DATA_BLOCK "TCP_IP_Shuttle_DB_20"   // DB238
{ S7_Optimized_Access := 'TRUE' }
VERSION : 0.1
// stored: AutoNumber true, DBAccessibleFromOPCUA true, IsOnlyStoredInLoadMemory false, IsRetainMemResEnabled false, IsWriteProtectedInAS false, MemoryReserve 100
   VAR
      enable : Bool := TRUE;
      send : Bool;
      sendDataLength : UDInt := 0;
      receiveDataLength : UDInt := 16#FFFF_FFFF;
   END_VAR
   VAR RETAIN
      tcpConfig : "LCom_typeConfig";
   END_VAR
   VAR
      tcpDiagnostics { S7_SetPoint := 'True'} : "LCom_typeDiagnostics";
      sendBuffer { S7_SetPoint := 'True'} : Array[0..59] of Byte;
      SendBufferSize : UInt := 60;
      receiveBuffer : Array[0..27] of Byte;
      receiveBufferSize : UInt := 28;
      connected : Bool;
      sending : Bool;
      dataReceived : Bool;
      receivedDataLength : UDInt;
      busy : Bool;
      error : Bool;
      status : Word;
   END_VAR
BEGIN
   tcpConfig.connection.interfaceID := 65164;
   tcpConfig.connection.connectionID := 120;
   tcpConfig.connection.comService := 1;
   tcpConfig.connection.isClient := False;
   tcpConfig.connection.connectType := 1;
   tcpConfig.connection.localPort := 4020;
   tcpConfig.connection.partnerPort := 4020;
   tcpConfig.connection.partnerIP.ADDR[1] := 10;
   tcpConfig.connection.partnerIP.ADDR[2] := 0;
   tcpConfig.connection.partnerIP.ADDR[3] := 34;
   tcpConfig.connection.partnerIP.ADDR[4] := 230;
   tcpConfig.connection.acceptUnknownPartner := TRUE;
   tcpConfig.connection.lifeSignCycleTime := T#1s;
   // sendBuffer[0] : STX
   // sendBuffer[1] : Size
   // sendBuffer[2] : Type
   // sendBuffer[3] : Request ID 1
   // sendBuffer[4] : Request ID 2
   // sendBuffer[5] : PID 1
   // sendBuffer[6] : PID 2
   // sendBuffer[7] : PID 3
   // sendBuffer[8] : PID 4
   // sendBuffer[9] : DID 1
   // sendBuffer[10] : DID 2
   // sendBuffer[11] : DID 3
   // sendBuffer[12] : DID 4
   // sendBuffer[13] : Distance remaining 1
   // sendBuffer[14] : Distance remaining 2
   // sendBuffer[15] : X
   // sendBuffer[16] : X
   // sendBuffer[17] : X
   // sendBuffer[18] : X
   // sendBuffer[19] : Y
   // sendBuffer[20] : Y
   // sendBuffer[21] : Y
   // sendBuffer[22] : Y
   // sendBuffer[23] : Floor
   // sendBuffer[24] : Mode
   // sendBuffer[25] : State
   // sendBuffer[26] : Load State
   // sendBuffer[27] : E1
   // sendBuffer[28] : E1
   // sendBuffer[29] : E2
   // sendBuffer[30] : E2
   // sendBuffer[31] : E3
   // sendBuffer[32] : E3
   // sendBuffer[33] : E4
   // sendBuffer[34] : E4
   // sendBuffer[35] : E5
   // sendBuffer[36] : E5
   // sendBuffer[37] : E6
   // sendBuffer[38] : E6
   // sendBuffer[39] : I1
   // sendBuffer[40] : I1
   // sendBuffer[41] : Q1
   // sendBuffer[42] : Q1
   // sendBuffer[43] : Barcode 1
   // sendBuffer[44] : Barcode 2
   // sendBuffer[45] : Barcode 3
   // sendBuffer[46] : Barcode 4
   // sendBuffer[47] : Pallet Type
   // sendBuffer[48] : Energy Level
   // sendBuffer[49] : Battery Voltage
   // sendBuffer[50] : Battery Voltage
   // sendBuffer[51] : Paused
   // sendBuffer[52] : Last order 1
   // sendBuffer[53] : Last order 2
   // sendBuffer[54] : Current order 1
   // sendBuffer[55] : Current order 2
   // sendBuffer[56] : Last finished 1
   // sendBuffer[57] : Last Finished 2
   // sendBuffer[58] : CS
   // sendBuffer[59] : ETX
   // receiveBuffer[0] : STX
   // receiveBuffer[1] : Size (length of payload)
   // receiveBuffer[2] : Type
   // receiveBuffer[3] : Request ID 1
   // receiveBuffer[4] : Request ID 2
END_DATA_BLOCK

DATA_BLOCK "TCP_IP_Shuttle_DB_21"   // DB166
{ S7_Optimized_Access := 'TRUE' }
VERSION : 0.1
// stored: AutoNumber true, DBAccessibleFromOPCUA true, IsOnlyStoredInLoadMemory false, IsRetainMemResEnabled false, IsWriteProtectedInAS false, MemoryReserve 100
   VAR
      enable : Bool := TRUE;
      send : Bool;
      sendDataLength : UDInt := 0;
      receiveDataLength : UDInt := 16#FFFF_FFFF;
   END_VAR
   VAR RETAIN
      tcpConfig : "LCom_typeConfig";
   END_VAR
   VAR
      tcpDiagnostics { S7_SetPoint := 'True'} : "LCom_typeDiagnostics";
      sendBuffer { S7_SetPoint := 'True'} : Array[0..59] of Byte;
      SendBufferSize : UInt := 60;
      receiveBuffer : Array[0..27] of Byte;
      receiveBufferSize : UInt := 28;
      connected : Bool;
      sending : Bool;
      dataReceived : Bool;
      receivedDataLength : UDInt;
      busy : Bool;
      error : Bool;
      status : Word;
   END_VAR
BEGIN
   tcpConfig.connection.interfaceID := 65164;
   tcpConfig.connection.connectionID := 121;
   tcpConfig.connection.comService := 1;
   tcpConfig.connection.isClient := False;
   tcpConfig.connection.connectType := 1;
   tcpConfig.connection.localPort := 4021;
   tcpConfig.connection.partnerPort := 4021;
   tcpConfig.connection.partnerIP.ADDR[1] := 10;
   tcpConfig.connection.partnerIP.ADDR[2] := 0;
   tcpConfig.connection.partnerIP.ADDR[3] := 34;
   tcpConfig.connection.partnerIP.ADDR[4] := 231;
   tcpConfig.connection.acceptUnknownPartner := TRUE;
   tcpConfig.connection.lifeSignCycleTime := T#1s;
   // sendBuffer[0] : STX
   // sendBuffer[1] : Size
   // sendBuffer[2] : Type
   // sendBuffer[3] : Request ID 1
   // sendBuffer[4] : Request ID 2
   // sendBuffer[5] : PID 1
   // sendBuffer[6] : PID 2
   // sendBuffer[7] : PID 3
   // sendBuffer[8] : PID 4
   // sendBuffer[9] : DID 1
   // sendBuffer[10] : DID 2
   // sendBuffer[11] : DID 3
   // sendBuffer[12] : DID 4
   // sendBuffer[13] : Distance remaining 1
   // sendBuffer[14] : Distance remaining 2
   // sendBuffer[15] : X
   // sendBuffer[16] : X
   // sendBuffer[17] : X
   // sendBuffer[18] : X
   // sendBuffer[19] : Y
   // sendBuffer[20] : Y
   // sendBuffer[21] : Y
   // sendBuffer[22] : Y
   // sendBuffer[23] : Floor
   // sendBuffer[24] : Mode
   // sendBuffer[25] : State
   // sendBuffer[26] : Load State
   // sendBuffer[27] : E1
   // sendBuffer[28] : E1
   // sendBuffer[29] : E2
   // sendBuffer[30] : E2
   // sendBuffer[31] : E3
   // sendBuffer[32] : E3
   // sendBuffer[33] : E4
   // sendBuffer[34] : E4
   // sendBuffer[35] : E5
   // sendBuffer[36] : E5
   // sendBuffer[37] : E6
   // sendBuffer[38] : E6
   // sendBuffer[39] : I1
   // sendBuffer[40] : I1
   // sendBuffer[41] : Q1
   // sendBuffer[42] : Q1
   // sendBuffer[43] : Barcode 1
   // sendBuffer[44] : Barcode 2
   // sendBuffer[45] : Barcode 3
   // sendBuffer[46] : Barcode 4
   // sendBuffer[47] : Pallet Type
   // sendBuffer[48] : Energy Level
   // sendBuffer[49] : Battery Voltage
   // sendBuffer[50] : Battery Voltage
   // sendBuffer[51] : Paused
   // sendBuffer[52] : Last order 1
   // sendBuffer[53] : Last order 2
   // sendBuffer[54] : Current order 1
   // sendBuffer[55] : Current order 2
   // sendBuffer[56] : Last finished 1
   // sendBuffer[57] : Last Finished 2
   // sendBuffer[58] : CS
   // sendBuffer[59] : ETX
   // receiveBuffer[0] : STX
   // receiveBuffer[1] : Size (length of payload)
   // receiveBuffer[2] : Type
   // receiveBuffer[3] : Request ID 1
   // receiveBuffer[4] : Request ID 2
END_DATA_BLOCK

DATA_BLOCK "TCP_IP_Shuttle_DB_22"   // DB241
{ S7_Optimized_Access := 'TRUE' }
VERSION : 0.1
// stored: AutoNumber true, DBAccessibleFromOPCUA true, IsOnlyStoredInLoadMemory false, IsRetainMemResEnabled false, IsWriteProtectedInAS false, MemoryReserve 100
   VAR
      enable : Bool := TRUE;
      send : Bool;
      sendDataLength : UDInt := 0;
      receiveDataLength : UDInt := 16#FFFF_FFFF;
   END_VAR
   VAR RETAIN
      tcpConfig : "LCom_typeConfig";
   END_VAR
   VAR
      tcpDiagnostics { S7_SetPoint := 'True'} : "LCom_typeDiagnostics";
      sendBuffer { S7_SetPoint := 'True'} : Array[0..59] of Byte;
      SendBufferSize : UInt := 60;
      receiveBuffer : Array[0..27] of Byte;
      receiveBufferSize : UInt := 28;
      connected : Bool;
      sending : Bool;
      dataReceived : Bool;
      receivedDataLength : UDInt;
      busy : Bool;
      error : Bool;
      status : Word;
   END_VAR
BEGIN
   tcpConfig.connection.interfaceID := 65164;
   tcpConfig.connection.connectionID := 122;
   tcpConfig.connection.comService := 1;
   tcpConfig.connection.isClient := False;
   tcpConfig.connection.connectType := 1;
   tcpConfig.connection.localPort := 4022;
   tcpConfig.connection.partnerPort := 4022;
   tcpConfig.connection.partnerIP.ADDR[1] := 10;
   tcpConfig.connection.partnerIP.ADDR[2] := 0;
   tcpConfig.connection.partnerIP.ADDR[3] := 34;
   tcpConfig.connection.partnerIP.ADDR[4] := 232;
   tcpConfig.connection.acceptUnknownPartner := TRUE;
   tcpConfig.connection.lifeSignCycleTime := T#1s;
   // sendBuffer[0] : STX
   // sendBuffer[1] : Size
   // sendBuffer[2] : Type
   // sendBuffer[3] : Request ID 1
   // sendBuffer[4] : Request ID 2
   // sendBuffer[5] : PID 1
   // sendBuffer[6] : PID 2
   // sendBuffer[7] : PID 3
   // sendBuffer[8] : PID 4
   // sendBuffer[9] : DID 1
   // sendBuffer[10] : DID 2
   // sendBuffer[11] : DID 3
   // sendBuffer[12] : DID 4
   // sendBuffer[13] : Distance remaining 1
   // sendBuffer[14] : Distance remaining 2
   // sendBuffer[15] : X
   // sendBuffer[16] : X
   // sendBuffer[17] : X
   // sendBuffer[18] : X
   // sendBuffer[19] : Y
   // sendBuffer[20] : Y
   // sendBuffer[21] : Y
   // sendBuffer[22] : Y
   // sendBuffer[23] : Floor
   // sendBuffer[24] : Mode
   // sendBuffer[25] : State
   // sendBuffer[26] : Load State
   // sendBuffer[27] : E1
   // sendBuffer[28] : E1
   // sendBuffer[29] : E2
   // sendBuffer[30] : E2
   // sendBuffer[31] : E3
   // sendBuffer[32] : E3
   // sendBuffer[33] : E4
   // sendBuffer[34] : E4
   // sendBuffer[35] : E5
   // sendBuffer[36] : E5
   // sendBuffer[37] : E6
   // sendBuffer[38] : E6
   // sendBuffer[39] : I1
   // sendBuffer[40] : I1
   // sendBuffer[41] : Q1
   // sendBuffer[42] : Q1
   // sendBuffer[43] : Barcode 1
   // sendBuffer[44] : Barcode 2
   // sendBuffer[45] : Barcode 3
   // sendBuffer[46] : Barcode 4
   // sendBuffer[47] : Pallet Type
   // sendBuffer[48] : Energy Level
   // sendBuffer[49] : Battery Voltage
   // sendBuffer[50] : Battery Voltage
   // sendBuffer[51] : Paused
   // sendBuffer[52] : Last order 1
   // sendBuffer[53] : Last order 2
   // sendBuffer[54] : Current order 1
   // sendBuffer[55] : Current order 2
   // sendBuffer[56] : Last finished 1
   // sendBuffer[57] : Last Finished 2
   // sendBuffer[58] : CS
   // sendBuffer[59] : ETX
   // receiveBuffer[0] : STX
   // receiveBuffer[1] : Size (length of payload)
   // receiveBuffer[2] : Type
   // receiveBuffer[3] : Request ID 1
   // receiveBuffer[4] : Request ID 2
END_DATA_BLOCK

DATA_BLOCK "TCP_IP_Shuttle_DB_23"   // DB382
{ S7_Optimized_Access := 'TRUE' }
VERSION : 0.1
// stored: AutoNumber true, DBAccessibleFromOPCUA true, IsOnlyStoredInLoadMemory false, IsRetainMemResEnabled false, IsWriteProtectedInAS false, MemoryReserve 100
   VAR
      enable : Bool := TRUE;
      send : Bool;
      sendDataLength : UDInt := 0;
      receiveDataLength : UDInt := 16#FFFF_FFFF;
   END_VAR
   VAR RETAIN
      tcpConfig : "LCom_typeConfig";
   END_VAR
   VAR
      tcpDiagnostics { S7_SetPoint := 'True'} : "LCom_typeDiagnostics";
      sendBuffer { S7_SetPoint := 'True'} : Array[0..59] of Byte;
      SendBufferSize : UInt := 60;
      receiveBuffer : Array[0..27] of Byte;
      receiveBufferSize : UInt := 28;
      connected : Bool;
      sending : Bool;
      dataReceived : Bool;
      receivedDataLength : UDInt;
      busy : Bool;
      error : Bool;
      status : Word;
   END_VAR
BEGIN
   tcpConfig.connection.interfaceID := 65164;
   tcpConfig.connection.connectionID := 123;
   tcpConfig.connection.comService := 1;
   tcpConfig.connection.isClient := False;
   tcpConfig.connection.connectType := 1;
   tcpConfig.connection.localPort := 4023;
   tcpConfig.connection.partnerPort := 4023;
   tcpConfig.connection.partnerIP.ADDR[1] := 10;
   tcpConfig.connection.partnerIP.ADDR[2] := 0;
   tcpConfig.connection.partnerIP.ADDR[3] := 34;
   tcpConfig.connection.partnerIP.ADDR[4] := 233;
   tcpConfig.connection.acceptUnknownPartner := TRUE;
   tcpConfig.connection.lifeSignCycleTime := T#1s;
   // sendBuffer[0] : STX
   // sendBuffer[1] : Size
   // sendBuffer[2] : Type
   // sendBuffer[3] : Request ID 1
   // sendBuffer[4] : Request ID 2
   // sendBuffer[5] : PID 1
   // sendBuffer[6] : PID 2
   // sendBuffer[7] : PID 3
   // sendBuffer[8] : PID 4
   // sendBuffer[9] : DID 1
   // sendBuffer[10] : DID 2
   // sendBuffer[11] : DID 3
   // sendBuffer[12] : DID 4
   // sendBuffer[13] : Distance remaining 1
   // sendBuffer[14] : Distance remaining 2
   // sendBuffer[15] : X
   // sendBuffer[16] : X
   // sendBuffer[17] : X
   // sendBuffer[18] : X
   // sendBuffer[19] : Y
   // sendBuffer[20] : Y
   // sendBuffer[21] : Y
   // sendBuffer[22] : Y
   // sendBuffer[23] : Floor
   // sendBuffer[24] : Mode
   // sendBuffer[25] : State
   // sendBuffer[26] : Load State
   // sendBuffer[27] : E1
   // sendBuffer[28] : E1
   // sendBuffer[29] : E2
   // sendBuffer[30] : E2
   // sendBuffer[31] : E3
   // sendBuffer[32] : E3
   // sendBuffer[33] : E4
   // sendBuffer[34] : E4
   // sendBuffer[35] : E5
   // sendBuffer[36] : E5
   // sendBuffer[37] : E6
   // sendBuffer[38] : E6
   // sendBuffer[39] : I1
   // sendBuffer[40] : I1
   // sendBuffer[41] : Q1
   // sendBuffer[42] : Q1
   // sendBuffer[43] : Barcode 1
   // sendBuffer[44] : Barcode 2
   // sendBuffer[45] : Barcode 3
   // sendBuffer[46] : Barcode 4
   // sendBuffer[47] : Pallet Type
   // sendBuffer[48] : Energy Level
   // sendBuffer[49] : Battery Voltage
   // sendBuffer[50] : Battery Voltage
   // sendBuffer[51] : Paused
   // sendBuffer[52] : Last order 1
   // sendBuffer[53] : Last order 2
   // sendBuffer[54] : Current order 1
   // sendBuffer[55] : Current order 2
   // sendBuffer[56] : Last finished 1
   // sendBuffer[57] : Last Finished 2
   // sendBuffer[58] : CS
   // sendBuffer[59] : ETX
   // receiveBuffer[0] : STX
   // receiveBuffer[1] : Size (length of payload)
   // receiveBuffer[2] : Type
   // receiveBuffer[3] : Request ID 1
   // receiveBuffer[4] : Request ID 2
END_DATA_BLOCK

DATA_BLOCK "TCP_IP_Shuttle_DB_3"   // DB388
{ S7_Optimized_Access := 'TRUE' }
VERSION : 0.1
// stored: AutoNumber true, DBAccessibleFromOPCUA true, IsOnlyStoredInLoadMemory false, IsRetainMemResEnabled false, IsWriteProtectedInAS false, MemoryReserve 100
   VAR
      enable : Bool := TRUE;
      send : Bool;
      sendDataLength : UDInt := 0;
      receiveDataLength : UDInt := 16#FFFF_FFFF;
   END_VAR
   VAR RETAIN
      tcpConfig : "LCom_typeConfig";
   END_VAR
   VAR
      tcpDiagnostics { S7_SetPoint := 'True'} : "LCom_typeDiagnostics";
      sendBuffer { S7_SetPoint := 'True'} : Array[0..59] of Byte;
      SendBufferSize : UInt := 60;
      receiveBuffer : Array[0..27] of Byte;
      receiveBufferSize : UInt := 28;
      connected : Bool;
      sending : Bool;
      dataReceived : Bool;
      receivedDataLength : UDInt;
      busy : Bool;
      error : Bool;
      status : Word;
   END_VAR
BEGIN
   tcpConfig.connection.interfaceID := 65164;
   tcpConfig.connection.connectionID := 103;
   tcpConfig.connection.comService := 1;
   tcpConfig.connection.isClient := False;
   tcpConfig.connection.connectType := 1;
   tcpConfig.connection.localPort := 4003;
   tcpConfig.connection.partnerPort := 4003;
   tcpConfig.connection.partnerIP.ADDR[1] := 10;
   tcpConfig.connection.partnerIP.ADDR[2] := 0;
   tcpConfig.connection.partnerIP.ADDR[3] := 34;
   tcpConfig.connection.partnerIP.ADDR[4] := 213;
   tcpConfig.connection.acceptUnknownPartner := TRUE;
   tcpConfig.connection.lifeSignCycleTime := T#1s;
   // sendBuffer[0] : STX
   // sendBuffer[1] : Size
   // sendBuffer[2] : Type
   // sendBuffer[3] : Request ID 1
   // sendBuffer[4] : Request ID 2
   // sendBuffer[5] : PID 1
   // sendBuffer[6] : PID 2
   // sendBuffer[7] : PID 3
   // sendBuffer[8] : PID 4
   // sendBuffer[9] : DID 1
   // sendBuffer[10] : DID 2
   // sendBuffer[11] : DID 3
   // sendBuffer[12] : DID 4
   // sendBuffer[13] : Distance remaining 1
   // sendBuffer[14] : Distance remaining 2
   // sendBuffer[15] : X
   // sendBuffer[16] : X
   // sendBuffer[17] : X
   // sendBuffer[18] : X
   // sendBuffer[19] : Y
   // sendBuffer[20] : Y
   // sendBuffer[21] : Y
   // sendBuffer[22] : Y
   // sendBuffer[23] : Floor
   // sendBuffer[24] : Mode
   // sendBuffer[25] : State
   // sendBuffer[26] : Load State
   // sendBuffer[27] : E1
   // sendBuffer[28] : E1
   // sendBuffer[29] : E2
   // sendBuffer[30] : E2
   // sendBuffer[31] : E3
   // sendBuffer[32] : E3
   // sendBuffer[33] : E4
   // sendBuffer[34] : E4
   // sendBuffer[35] : E5
   // sendBuffer[36] : E5
   // sendBuffer[37] : E6
   // sendBuffer[38] : E6
   // sendBuffer[39] : I1
   // sendBuffer[40] : I1
   // sendBuffer[41] : Q1
   // sendBuffer[42] : Q1
   // sendBuffer[43] : Barcode 1
   // sendBuffer[44] : Barcode 2
   // sendBuffer[45] : Barcode 3
   // sendBuffer[46] : Barcode 4
   // sendBuffer[47] : Pallet Type
   // sendBuffer[48] : Energy Level
   // sendBuffer[49] : Battery Voltage
   // sendBuffer[50] : Battery Voltage
   // sendBuffer[51] : Paused
   // sendBuffer[52] : Last order 1
   // sendBuffer[53] : Last order 2
   // sendBuffer[54] : Current order 1
   // sendBuffer[55] : Current order 2
   // sendBuffer[56] : Last finished 1
   // sendBuffer[57] : Last Finished 2
   // sendBuffer[58] : CS
   // sendBuffer[59] : ETX
   // receiveBuffer[0] : STX
   // receiveBuffer[1] : Size (length of payload)
   // receiveBuffer[2] : Type
   // receiveBuffer[3] : Request ID 1
   // receiveBuffer[4] : Request ID 2
END_DATA_BLOCK

DATA_BLOCK "TCP_IP_Shuttle_DB_4"   // DB375
{ S7_Optimized_Access := 'TRUE' }
VERSION : 0.1
// stored: AutoNumber true, DBAccessibleFromOPCUA true, IsOnlyStoredInLoadMemory false, IsRetainMemResEnabled false, IsWriteProtectedInAS false, MemoryReserve 100
   VAR
      enable : Bool := TRUE;
      send : Bool;
      sendDataLength : UDInt := 0;
      receiveDataLength : UDInt := 16#FFFF_FFFF;
   END_VAR
   VAR RETAIN
      tcpConfig : "LCom_typeConfig";
   END_VAR
   VAR
      tcpDiagnostics { S7_SetPoint := 'True'} : "LCom_typeDiagnostics";
      sendBuffer { S7_SetPoint := 'True'} : Array[0..59] of Byte;
      SendBufferSize : UInt := 60;
      receiveBuffer : Array[0..27] of Byte;
      receiveBufferSize : UInt := 28;
      connected : Bool;
      sending : Bool;
      dataReceived : Bool;
      receivedDataLength : UDInt;
      busy : Bool;
      error : Bool;
      status : Word;
   END_VAR
BEGIN
   tcpConfig.connection.interfaceID := 65164;
   tcpConfig.connection.connectionID := 104;
   tcpConfig.connection.comService := 1;
   tcpConfig.connection.isClient := False;
   tcpConfig.connection.connectType := 1;
   tcpConfig.connection.localPort := 4004;
   tcpConfig.connection.partnerPort := 4004;
   tcpConfig.connection.partnerIP.ADDR[1] := 10;
   tcpConfig.connection.partnerIP.ADDR[2] := 0;
   tcpConfig.connection.partnerIP.ADDR[3] := 34;
   tcpConfig.connection.partnerIP.ADDR[4] := 214;
   tcpConfig.connection.acceptUnknownPartner := TRUE;
   tcpConfig.connection.lifeSignCycleTime := T#1s;
   // sendBuffer[0] : STX
   // sendBuffer[1] : Size
   // sendBuffer[2] : Type
   // sendBuffer[3] : Request ID 1
   // sendBuffer[4] : Request ID 2
   // sendBuffer[5] : PID 1
   // sendBuffer[6] : PID 2
   // sendBuffer[7] : PID 3
   // sendBuffer[8] : PID 4
   // sendBuffer[9] : DID 1
   // sendBuffer[10] : DID 2
   // sendBuffer[11] : DID 3
   // sendBuffer[12] : DID 4
   // sendBuffer[13] : Distance remaining 1
   // sendBuffer[14] : Distance remaining 2
   // sendBuffer[15] : X
   // sendBuffer[16] : X
   // sendBuffer[17] : X
   // sendBuffer[18] : X
   // sendBuffer[19] : Y
   // sendBuffer[20] : Y
   // sendBuffer[21] : Y
   // sendBuffer[22] : Y
   // sendBuffer[23] : Floor
   // sendBuffer[24] : Mode
   // sendBuffer[25] : State
   // sendBuffer[26] : Load State
   // sendBuffer[27] : E1
   // sendBuffer[28] : E1
   // sendBuffer[29] : E2
   // sendBuffer[30] : E2
   // sendBuffer[31] : E3
   // sendBuffer[32] : E3
   // sendBuffer[33] : E4
   // sendBuffer[34] : E4
   // sendBuffer[35] : E5
   // sendBuffer[36] : E5
   // sendBuffer[37] : E6
   // sendBuffer[38] : E6
   // sendBuffer[39] : I1
   // sendBuffer[40] : I1
   // sendBuffer[41] : Q1
   // sendBuffer[42] : Q1
   // sendBuffer[43] : Barcode 1
   // sendBuffer[44] : Barcode 2
   // sendBuffer[45] : Barcode 3
   // sendBuffer[46] : Barcode 4
   // sendBuffer[47] : Pallet Type
   // sendBuffer[48] : Energy Level
   // sendBuffer[49] : Battery Voltage
   // sendBuffer[50] : Battery Voltage
   // sendBuffer[51] : Paused
   // sendBuffer[52] : Last order 1
   // sendBuffer[53] : Last order 2
   // sendBuffer[54] : Current order 1
   // sendBuffer[55] : Current order 2
   // sendBuffer[56] : Last finished 1
   // sendBuffer[57] : Last Finished 2
   // sendBuffer[58] : CS
   // sendBuffer[59] : ETX
   // receiveBuffer[0] : STX
   // receiveBuffer[1] : Size (length of payload)
   // receiveBuffer[2] : Type
   // receiveBuffer[3] : Request ID 1
   // receiveBuffer[4] : Request ID 2
END_DATA_BLOCK

DATA_BLOCK "TCP_IP_Shuttle_DB_5"   // DB376
{ S7_Optimized_Access := 'TRUE' }
VERSION : 0.1
// stored: AutoNumber true, DBAccessibleFromOPCUA true, IsOnlyStoredInLoadMemory false, IsRetainMemResEnabled false, IsWriteProtectedInAS false, MemoryReserve 100
   VAR
      enable : Bool := TRUE;
      send : Bool;
      sendDataLength : UDInt := 0;
      receiveDataLength : UDInt := 16#FFFF_FFFF;
   END_VAR
   VAR RETAIN
      tcpConfig : "LCom_typeConfig";
   END_VAR
   VAR
      tcpDiagnostics { S7_SetPoint := 'True'} : "LCom_typeDiagnostics";
      sendBuffer { S7_SetPoint := 'True'} : Array[0..59] of Byte;
      SendBufferSize : UInt := 60;
      receiveBuffer : Array[0..27] of Byte;
      receiveBufferSize : UInt := 28;
      connected : Bool;
      sending : Bool;
      dataReceived : Bool;
      receivedDataLength : UDInt;
      busy : Bool;
      error : Bool;
      status : Word;
   END_VAR
BEGIN
   tcpConfig.connection.interfaceID := 65164;
   tcpConfig.connection.connectionID := 105;
   tcpConfig.connection.comService := 1;
   tcpConfig.connection.isClient := False;
   tcpConfig.connection.connectType := 1;
   tcpConfig.connection.localPort := 4005;
   tcpConfig.connection.partnerPort := 4005;
   tcpConfig.connection.partnerIP.ADDR[1] := 10;
   tcpConfig.connection.partnerIP.ADDR[2] := 0;
   tcpConfig.connection.partnerIP.ADDR[3] := 34;
   tcpConfig.connection.partnerIP.ADDR[4] := 215;
   tcpConfig.connection.acceptUnknownPartner := TRUE;
   tcpConfig.connection.lifeSignCycleTime := T#1s;
   // sendBuffer[0] : STX
   // sendBuffer[1] : Size
   // sendBuffer[2] : Type
   // sendBuffer[3] : Request ID 1
   // sendBuffer[4] : Request ID 2
   // sendBuffer[5] : PID 1
   // sendBuffer[6] : PID 2
   // sendBuffer[7] : PID 3
   // sendBuffer[8] : PID 4
   // sendBuffer[9] : DID 1
   // sendBuffer[10] : DID 2
   // sendBuffer[11] : DID 3
   // sendBuffer[12] : DID 4
   // sendBuffer[13] : Distance remaining 1
   // sendBuffer[14] : Distance remaining 2
   // sendBuffer[15] : X
   // sendBuffer[16] : X
   // sendBuffer[17] : X
   // sendBuffer[18] : X
   // sendBuffer[19] : Y
   // sendBuffer[20] : Y
   // sendBuffer[21] : Y
   // sendBuffer[22] : Y
   // sendBuffer[23] : Floor
   // sendBuffer[24] : Mode
   // sendBuffer[25] : State
   // sendBuffer[26] : Load State
   // sendBuffer[27] : E1
   // sendBuffer[28] : E1
   // sendBuffer[29] : E2
   // sendBuffer[30] : E2
   // sendBuffer[31] : E3
   // sendBuffer[32] : E3
   // sendBuffer[33] : E4
   // sendBuffer[34] : E4
   // sendBuffer[35] : E5
   // sendBuffer[36] : E5
   // sendBuffer[37] : E6
   // sendBuffer[38] : E6
   // sendBuffer[39] : I1
   // sendBuffer[40] : I1
   // sendBuffer[41] : Q1
   // sendBuffer[42] : Q1
   // sendBuffer[43] : Barcode 1
   // sendBuffer[44] : Barcode 2
   // sendBuffer[45] : Barcode 3
   // sendBuffer[46] : Barcode 4
   // sendBuffer[47] : Pallet Type
   // sendBuffer[48] : Energy Level
   // sendBuffer[49] : Battery Voltage
   // sendBuffer[50] : Battery Voltage
   // sendBuffer[51] : Paused
   // sendBuffer[52] : Last order 1
   // sendBuffer[53] : Last order 2
   // sendBuffer[54] : Current order 1
   // sendBuffer[55] : Current order 2
   // sendBuffer[56] : Last finished 1
   // sendBuffer[57] : Last Finished 2
   // sendBuffer[58] : CS
   // sendBuffer[59] : ETX
   // receiveBuffer[0] : STX
   // receiveBuffer[1] : Size (length of payload)
   // receiveBuffer[2] : Type
   // receiveBuffer[3] : Request ID 1
   // receiveBuffer[4] : Request ID 2
END_DATA_BLOCK

DATA_BLOCK "TCP_IP_Shuttle_DB_6"   // DB377
{ S7_Optimized_Access := 'TRUE' }
VERSION : 0.1
// stored: AutoNumber true, DBAccessibleFromOPCUA true, IsOnlyStoredInLoadMemory false, IsRetainMemResEnabled false, IsWriteProtectedInAS false, MemoryReserve 100
   VAR
      enable : Bool := TRUE;
      send : Bool;
      sendDataLength : UDInt := 0;
      receiveDataLength : UDInt := 16#FFFF_FFFF;
   END_VAR
   VAR RETAIN
      tcpConfig : "LCom_typeConfig";
   END_VAR
   VAR
      tcpDiagnostics { S7_SetPoint := 'True'} : "LCom_typeDiagnostics";
      sendBuffer { S7_SetPoint := 'True'} : Array[0..59] of Byte;
      SendBufferSize : UInt := 60;
      receiveBuffer : Array[0..27] of Byte;
      receiveBufferSize : UInt := 28;
      connected : Bool;
      sending : Bool;
      dataReceived : Bool;
      receivedDataLength : UDInt;
      busy : Bool;
      error : Bool;
      status : Word;
   END_VAR
BEGIN
   tcpConfig.connection.interfaceID := 65164;
   tcpConfig.connection.connectionID := 106;
   tcpConfig.connection.comService := 1;
   tcpConfig.connection.isClient := False;
   tcpConfig.connection.connectType := 1;
   tcpConfig.connection.localPort := 4006;
   tcpConfig.connection.partnerPort := 4006;
   tcpConfig.connection.partnerIP.ADDR[1] := 10;
   tcpConfig.connection.partnerIP.ADDR[2] := 0;
   tcpConfig.connection.partnerIP.ADDR[3] := 34;
   tcpConfig.connection.partnerIP.ADDR[4] := 216;
   tcpConfig.connection.acceptUnknownPartner := TRUE;
   tcpConfig.connection.lifeSignCycleTime := T#1s;
   // sendBuffer[0] : STX
   // sendBuffer[1] : Size
   // sendBuffer[2] : Type
   // sendBuffer[3] : Request ID 1
   // sendBuffer[4] : Request ID 2
   // sendBuffer[5] : PID 1
   // sendBuffer[6] : PID 2
   // sendBuffer[7] : PID 3
   // sendBuffer[8] : PID 4
   // sendBuffer[9] : DID 1
   // sendBuffer[10] : DID 2
   // sendBuffer[11] : DID 3
   // sendBuffer[12] : DID 4
   // sendBuffer[13] : Distance remaining 1
   // sendBuffer[14] : Distance remaining 2
   // sendBuffer[15] : X
   // sendBuffer[16] : X
   // sendBuffer[17] : X
   // sendBuffer[18] : X
   // sendBuffer[19] : Y
   // sendBuffer[20] : Y
   // sendBuffer[21] : Y
   // sendBuffer[22] : Y
   // sendBuffer[23] : Floor
   // sendBuffer[24] : Mode
   // sendBuffer[25] : State
   // sendBuffer[26] : Load State
   // sendBuffer[27] : E1
   // sendBuffer[28] : E1
   // sendBuffer[29] : E2
   // sendBuffer[30] : E2
   // sendBuffer[31] : E3
   // sendBuffer[32] : E3
   // sendBuffer[33] : E4
   // sendBuffer[34] : E4
   // sendBuffer[35] : E5
   // sendBuffer[36] : E5
   // sendBuffer[37] : E6
   // sendBuffer[38] : E6
   // sendBuffer[39] : I1
   // sendBuffer[40] : I1
   // sendBuffer[41] : Q1
   // sendBuffer[42] : Q1
   // sendBuffer[43] : Barcode 1
   // sendBuffer[44] : Barcode 2
   // sendBuffer[45] : Barcode 3
   // sendBuffer[46] : Barcode 4
   // sendBuffer[47] : Pallet Type
   // sendBuffer[48] : Energy Level
   // sendBuffer[49] : Battery Voltage
   // sendBuffer[50] : Battery Voltage
   // sendBuffer[51] : Paused
   // sendBuffer[52] : Last order 1
   // sendBuffer[53] : Last order 2
   // sendBuffer[54] : Current order 1
   // sendBuffer[55] : Current order 2
   // sendBuffer[56] : Last finished 1
   // sendBuffer[57] : Last Finished 2
   // sendBuffer[58] : CS
   // sendBuffer[59] : ETX
   // receiveBuffer[0] : STX
   // receiveBuffer[1] : Size (length of payload)
   // receiveBuffer[2] : Type
   // receiveBuffer[3] : Request ID 1
   // receiveBuffer[4] : Request ID 2
END_DATA_BLOCK

DATA_BLOCK "TCP_IP_Shuttle_DB_7"   // DB374
{ S7_Optimized_Access := 'TRUE' }
VERSION : 0.1
// stored: AutoNumber true, DBAccessibleFromOPCUA true, IsOnlyStoredInLoadMemory false, IsRetainMemResEnabled false, IsWriteProtectedInAS false, MemoryReserve 100
   VAR
      enable : Bool := TRUE;
      send : Bool;
      sendDataLength : UDInt := 0;
      receiveDataLength : UDInt := 16#FFFF_FFFF;
   END_VAR
   VAR RETAIN
      tcpConfig : "LCom_typeConfig";
   END_VAR
   VAR
      tcpDiagnostics { S7_SetPoint := 'True'} : "LCom_typeDiagnostics";
      sendBuffer { S7_SetPoint := 'True'} : Array[0..59] of Byte;
      SendBufferSize : UInt := 60;
      receiveBuffer : Array[0..27] of Byte;
      receiveBufferSize : UInt := 28;
      connected : Bool;
      sending : Bool;
      dataReceived : Bool;
      receivedDataLength : UDInt;
      busy : Bool;
      error : Bool;
      status : Word;
   END_VAR
BEGIN
   tcpConfig.connection.interfaceID := 65164;
   tcpConfig.connection.connectionID := 107;
   tcpConfig.connection.comService := 1;
   tcpConfig.connection.isClient := False;
   tcpConfig.connection.connectType := 1;
   tcpConfig.connection.localPort := 4007;
   tcpConfig.connection.partnerPort := 4007;
   tcpConfig.connection.partnerIP.ADDR[1] := 10;
   tcpConfig.connection.partnerIP.ADDR[2] := 0;
   tcpConfig.connection.partnerIP.ADDR[3] := 34;
   tcpConfig.connection.partnerIP.ADDR[4] := 217;
   tcpConfig.connection.acceptUnknownPartner := TRUE;
   tcpConfig.connection.lifeSignCycleTime := T#1s;
   // sendBuffer[0] : STX
   // sendBuffer[1] : Size
   // sendBuffer[2] : Type
   // sendBuffer[3] : Request ID 1
   // sendBuffer[4] : Request ID 2
   // sendBuffer[5] : PID 1
   // sendBuffer[6] : PID 2
   // sendBuffer[7] : PID 3
   // sendBuffer[8] : PID 4
   // sendBuffer[9] : DID 1
   // sendBuffer[10] : DID 2
   // sendBuffer[11] : DID 3
   // sendBuffer[12] : DID 4
   // sendBuffer[13] : Distance remaining 1
   // sendBuffer[14] : Distance remaining 2
   // sendBuffer[15] : X
   // sendBuffer[16] : X
   // sendBuffer[17] : X
   // sendBuffer[18] : X
   // sendBuffer[19] : Y
   // sendBuffer[20] : Y
   // sendBuffer[21] : Y
   // sendBuffer[22] : Y
   // sendBuffer[23] : Floor
   // sendBuffer[24] : Mode
   // sendBuffer[25] : State
   // sendBuffer[26] : Load State
   // sendBuffer[27] : E1
   // sendBuffer[28] : E1
   // sendBuffer[29] : E2
   // sendBuffer[30] : E2
   // sendBuffer[31] : E3
   // sendBuffer[32] : E3
   // sendBuffer[33] : E4
   // sendBuffer[34] : E4
   // sendBuffer[35] : E5
   // sendBuffer[36] : E5
   // sendBuffer[37] : E6
   // sendBuffer[38] : E6
   // sendBuffer[39] : I1
   // sendBuffer[40] : I1
   // sendBuffer[41] : Q1
   // sendBuffer[42] : Q1
   // sendBuffer[43] : Barcode 1
   // sendBuffer[44] : Barcode 2
   // sendBuffer[45] : Barcode 3
   // sendBuffer[46] : Barcode 4
   // sendBuffer[47] : Pallet Type
   // sendBuffer[48] : Energy Level
   // sendBuffer[49] : Battery Voltage
   // sendBuffer[50] : Battery Voltage
   // sendBuffer[51] : Paused
   // sendBuffer[52] : Last order 1
   // sendBuffer[53] : Last order 2
   // sendBuffer[54] : Current order 1
   // sendBuffer[55] : Current order 2
   // sendBuffer[56] : Last finished 1
   // sendBuffer[57] : Last Finished 2
   // sendBuffer[58] : CS
   // sendBuffer[59] : ETX
   // receiveBuffer[0] : STX
   // receiveBuffer[1] : Size (length of payload)
   // receiveBuffer[2] : Type
   // receiveBuffer[3] : Request ID 1
   // receiveBuffer[4] : Request ID 2
END_DATA_BLOCK

DATA_BLOCK "TCP_IP_Shuttle_DB_8"   // DB380
{ S7_Optimized_Access := 'TRUE' }
VERSION : 0.1
// stored: AutoNumber true, DBAccessibleFromOPCUA true, IsOnlyStoredInLoadMemory false, IsRetainMemResEnabled false, IsWriteProtectedInAS false, MemoryReserve 100
   VAR
      enable : Bool := TRUE;
      send : Bool;
      sendDataLength : UDInt := 0;
      receiveDataLength : UDInt := 16#FFFF_FFFF;
   END_VAR
   VAR RETAIN
      tcpConfig : "LCom_typeConfig";
   END_VAR
   VAR
      tcpDiagnostics { S7_SetPoint := 'True'} : "LCom_typeDiagnostics";
      sendBuffer { S7_SetPoint := 'True'} : Array[0..59] of Byte;
      SendBufferSize : UInt := 60;
      receiveBuffer : Array[0..27] of Byte;
      receiveBufferSize : UInt := 28;
      connected : Bool;
      sending : Bool;
      dataReceived : Bool;
      receivedDataLength : UDInt;
      busy : Bool;
      error : Bool;
      status : Word;
   END_VAR
BEGIN
   tcpConfig.connection.interfaceID := 65164;
   tcpConfig.connection.connectionID := 108;
   tcpConfig.connection.comService := 1;
   tcpConfig.connection.isClient := False;
   tcpConfig.connection.connectType := 1;
   tcpConfig.connection.localPort := 4008;
   tcpConfig.connection.partnerPort := 4008;
   tcpConfig.connection.partnerIP.ADDR[1] := 10;
   tcpConfig.connection.partnerIP.ADDR[2] := 0;
   tcpConfig.connection.partnerIP.ADDR[3] := 34;
   tcpConfig.connection.partnerIP.ADDR[4] := 218;
   tcpConfig.connection.acceptUnknownPartner := TRUE;
   tcpConfig.connection.lifeSignCycleTime := T#1s;
   // sendBuffer[0] : STX
   // sendBuffer[1] : Size
   // sendBuffer[2] : Type
   // sendBuffer[3] : Request ID 1
   // sendBuffer[4] : Request ID 2
   // sendBuffer[5] : PID 1
   // sendBuffer[6] : PID 2
   // sendBuffer[7] : PID 3
   // sendBuffer[8] : PID 4
   // sendBuffer[9] : DID 1
   // sendBuffer[10] : DID 2
   // sendBuffer[11] : DID 3
   // sendBuffer[12] : DID 4
   // sendBuffer[13] : Distance remaining 1
   // sendBuffer[14] : Distance remaining 2
   // sendBuffer[15] : X
   // sendBuffer[16] : X
   // sendBuffer[17] : X
   // sendBuffer[18] : X
   // sendBuffer[19] : Y
   // sendBuffer[20] : Y
   // sendBuffer[21] : Y
   // sendBuffer[22] : Y
   // sendBuffer[23] : Floor
   // sendBuffer[24] : Mode
   // sendBuffer[25] : State
   // sendBuffer[26] : Load State
   // sendBuffer[27] : E1
   // sendBuffer[28] : E1
   // sendBuffer[29] : E2
   // sendBuffer[30] : E2
   // sendBuffer[31] : E3
   // sendBuffer[32] : E3
   // sendBuffer[33] : E4
   // sendBuffer[34] : E4
   // sendBuffer[35] : E5
   // sendBuffer[36] : E5
   // sendBuffer[37] : E6
   // sendBuffer[38] : E6
   // sendBuffer[39] : I1
   // sendBuffer[40] : I1
   // sendBuffer[41] : Q1
   // sendBuffer[42] : Q1
   // sendBuffer[43] : Barcode 1
   // sendBuffer[44] : Barcode 2
   // sendBuffer[45] : Barcode 3
   // sendBuffer[46] : Barcode 4
   // sendBuffer[47] : Pallet Type
   // sendBuffer[48] : Energy Level
   // sendBuffer[49] : Battery Voltage
   // sendBuffer[50] : Battery Voltage
   // sendBuffer[51] : Paused
   // sendBuffer[52] : Last order 1
   // sendBuffer[53] : Last order 2
   // sendBuffer[54] : Current order 1
   // sendBuffer[55] : Current order 2
   // sendBuffer[56] : Last finished 1
   // sendBuffer[57] : Last Finished 2
   // sendBuffer[58] : CS
   // sendBuffer[59] : ETX
   // receiveBuffer[0] : STX
   // receiveBuffer[1] : Size (length of payload)
   // receiveBuffer[2] : Type
   // receiveBuffer[3] : Request ID 1
   // receiveBuffer[4] : Request ID 2
END_DATA_BLOCK

DATA_BLOCK "TCP_IP_Shuttle_DB_9"   // DB383
{ S7_Optimized_Access := 'TRUE' }
VERSION : 0.1
// stored: AutoNumber true, DBAccessibleFromOPCUA true, IsOnlyStoredInLoadMemory false, IsRetainMemResEnabled false, IsWriteProtectedInAS false, MemoryReserve 100
   VAR
      enable : Bool := TRUE;
      send : Bool;
      sendDataLength : UDInt := 0;
      receiveDataLength : UDInt := 16#FFFF_FFFF;
   END_VAR
   VAR RETAIN
      tcpConfig : "LCom_typeConfig";
   END_VAR
   VAR
      tcpDiagnostics { S7_SetPoint := 'True'} : "LCom_typeDiagnostics";
      sendBuffer { S7_SetPoint := 'True'} : Array[0..59] of Byte;
      SendBufferSize : UInt := 60;
      receiveBuffer : Array[0..27] of Byte;
      receiveBufferSize : UInt := 28;
      connected : Bool;
      sending : Bool;
      dataReceived : Bool;
      receivedDataLength : UDInt;
      busy : Bool;
      error : Bool;
      status : Word;
   END_VAR
BEGIN
   tcpConfig.connection.interfaceID := 65164;
   tcpConfig.connection.connectionID := 109;
   tcpConfig.connection.comService := 1;
   tcpConfig.connection.isClient := False;
   tcpConfig.connection.connectType := 1;
   tcpConfig.connection.localPort := 4009;
   tcpConfig.connection.partnerPort := 4009;
   tcpConfig.connection.partnerIP.ADDR[1] := 10;
   tcpConfig.connection.partnerIP.ADDR[2] := 0;
   tcpConfig.connection.partnerIP.ADDR[3] := 34;
   tcpConfig.connection.partnerIP.ADDR[4] := 219;
   tcpConfig.connection.acceptUnknownPartner := TRUE;
   tcpConfig.connection.lifeSignCycleTime := T#1s;
   // sendBuffer[0] : STX
   // sendBuffer[1] : Size
   // sendBuffer[2] : Type
   // sendBuffer[3] : Request ID 1
   // sendBuffer[4] : Request ID 2
   // sendBuffer[5] : PID 1
   // sendBuffer[6] : PID 2
   // sendBuffer[7] : PID 3
   // sendBuffer[8] : PID 4
   // sendBuffer[9] : DID 1
   // sendBuffer[10] : DID 2
   // sendBuffer[11] : DID 3
   // sendBuffer[12] : DID 4
   // sendBuffer[13] : Distance remaining 1
   // sendBuffer[14] : Distance remaining 2
   // sendBuffer[15] : X
   // sendBuffer[16] : X
   // sendBuffer[17] : X
   // sendBuffer[18] : X
   // sendBuffer[19] : Y
   // sendBuffer[20] : Y
   // sendBuffer[21] : Y
   // sendBuffer[22] : Y
   // sendBuffer[23] : Floor
   // sendBuffer[24] : Mode
   // sendBuffer[25] : State
   // sendBuffer[26] : Load State
   // sendBuffer[27] : E1
   // sendBuffer[28] : E1
   // sendBuffer[29] : E2
   // sendBuffer[30] : E2
   // sendBuffer[31] : E3
   // sendBuffer[32] : E3
   // sendBuffer[33] : E4
   // sendBuffer[34] : E4
   // sendBuffer[35] : E5
   // sendBuffer[36] : E5
   // sendBuffer[37] : E6
   // sendBuffer[38] : E6
   // sendBuffer[39] : I1
   // sendBuffer[40] : I1
   // sendBuffer[41] : Q1
   // sendBuffer[42] : Q1
   // sendBuffer[43] : Barcode 1
   // sendBuffer[44] : Barcode 2
   // sendBuffer[45] : Barcode 3
   // sendBuffer[46] : Barcode 4
   // sendBuffer[47] : Pallet Type
   // sendBuffer[48] : Energy Level
   // sendBuffer[49] : Battery Voltage
   // sendBuffer[50] : Battery Voltage
   // sendBuffer[51] : Paused
   // sendBuffer[52] : Last order 1
   // sendBuffer[53] : Last order 2
   // sendBuffer[54] : Current order 1
   // sendBuffer[55] : Current order 2
   // sendBuffer[56] : Last finished 1
   // sendBuffer[57] : Last Finished 2
   // sendBuffer[58] : CS
   // sendBuffer[59] : ETX
   // receiveBuffer[0] : STX
   // receiveBuffer[1] : Size (length of payload)
   // receiveBuffer[2] : Type
   // receiveBuffer[3] : Request ID 1
   // receiveBuffer[4] : Request ID 2
END_DATA_BLOCK

DATA_BLOCK "Time"   // DB135
{ S7_Optimized_Access := 'TRUE' }
VERSION : 0.1
// stored: AutoNumber true, DBAccessibleFromOPCUA true, IsOnlyStoredInLoadMemory false, IsRetainMemResEnabled false, IsWriteProtectedInAS false, MemoryReserve 100
   VAR
      CurrentLocalTime : String := '06/10/2022 09:04:28';
      CurrentDTL : DTL := DTL#2022-06-10-09:04:28.050899826;
      PC_HeartBeat : Word := 16#6E87;
      PLC_HeartBeat : Word := 16#B1AA;
   END_VAR
BEGIN
END_DATA_BLOCK

DATA_BLOCK "VTD_HMI"   // DB57
{ S7_Optimized_Access := 'TRUE' }
VERSION : 0.1
// stored: AutoNumber true, DBAccessibleFromOPCUA true, IsOnlyStoredInLoadMemory false, IsRetainMemResEnabled false, IsWriteProtectedInAS false, MemoryReserve 100
   VAR
      Start_InBarcodeStation : Array[1..5] of Bool;
      Move_To_Level : Array[1..5] of UInt;
      Mode_Change : Array[1..5] of UInt;
      Manual_Down : Array[1..5] of Bool;
      Pallet_Type : Array[1..5] of UInt;
      Manual_Up : Array[1..5] of Bool;
      Task_ID : Array[1..5] of UInt;
      Reset : Array[1..5] of Bool;
      Enable : Array[1..5] of Bool;
      Progress : Array[1..5] of Int;
      Stop : Array[1..5] of Bool;
      Manual_DP_Extend : Array[1..5] of Bool;
      Manual_DP_Retract : Array[1..5] of Bool;
      ID : Array[1..5] of UInt;
      Cnv_Occupied : Array[1..5] of Bool;
      Motor_Status : Array[1..5] of UInt;
      ID_OLD : Array[1..5] of UInt;
      LE_Error : Array[1..5] of Bool;
      Mode : Array[1..5] of UInt;
      Encoder_Delta : Array[1..5] of Real;
      Warning : Array[1..5] of Bool;
      Current_Level : Array[1..5] of UInt;
      Error : Array[1..5] of Bool;
      Current_Task_ID : Array[1..5] of UInt;
      Pallet_Loaded : Array[1..5] of UInt;
      Stopped : Array[1..5] of Bool;
      SM_State : Array[1..5] of UInt;
      Shuttle_Loaded : Array[1..5] of UInt;
      DP_State : Array[1..5] of UInt;
      AE : Array[1..5] of Real;
      Docked : Array[1..5] of Bool;
      AE_Error : Array[1..5] of Bool;
      Enabled : Array[1..5] of Bool;
      Current_Task_Type : Array[1..5] of UInt;
      Running : Array[1..5] of Bool;
      LE : Array[1..5] of Real;
      Motor_Actual_Speed : Array[1..5] of UInt;
      Motor_SetPoint : Array[1..5] of UInt;
      Motor_Actual_Current : Array[1..5] of Real;
      Motor_Ready : Array[1..5] of Bool;
      "Chain Slack 1" : Array[1..5] of Bool;
      "Chain Slack 3" : Array[1..5] of Bool;
      "Chain Slack 2" : Array[1..5] of Bool;
      "Chain Slack 4" : Array[1..5] of Bool;
      Safety_OK : Array[1..5] of Bool;
      Moving_To_Level : Array[1..5] of UInt;
      Speed_mm_s : Array[1..5] of Real;
      Level_Below_Extractor : Array[1..5] of UInt;
      Actual_Torque : Array[1..5] of UInt;
      DP1_Retracted : Array[1..5] of Bool;
      DP2_Extended : Array[1..5] of Bool;
      Upper_Overtravel : Array[1..5] of Bool;
      DP1_Extended : Array[1..5] of Bool;
      DP2_Retracted : Array[1..5] of Bool;
      Lower_Overtravel : Array[1..5] of Bool;
      Level_Detect1 : Array[1..5] of Bool;
      Lower_Limit : Array[1..5] of Bool;
      Ultimate_Creep : Array[1..5] of Bool;
      Upper_Limet : Array[1..5] of Bool;
      Level_Detect2 : Array[1..5] of Bool;
      Ultimate_Slow : Array[1..5] of Bool;
      Charge_VTD_Commands : Array[1..5] of Bool;
      LE_Bypass : Array[1..5] of Bool;
      Charge_VTD : Array[1..5] of Bool;
   END_VAR
BEGIN
END_DATA_BLOCK

ORGANIZATION_BLOCK "Main"   // OB1, LAD, ProgramCycle
TITLE = "Main Program Sweep (Cycle)"
{ S7_Optimized_Access := 'TRUE' }
VERSION : 0.1
// stored: AutoNumber true, IsIECCheckEnabled false, SetENOAutomatically false
   VAR_INPUT
      Initial_Call : Bool;   // Initial call of this OB
      Remanence : Bool;   // =True, if remanent data are available
   END_VAR
   VAR_TEMP
      Fault_Handshake_Infeed_1 : Bool;
      Fault_Handshake_Outfeed_1 : Bool;
      Fault_Handshake_Infeed_2 : Bool;
      Fault_Handshake_Infeed_3 : Bool;
      Fault_Handshake_Outfeed_2 : Bool;
      Fault_Handshake_Outfeed_3 : Bool;
   END_VAR
   VAR_TEMP   // added for the SCL form of the ladder/FBD networks
      _w1 : Bool;
      _w2 : Bool;
      _w3 : Bool;
      _w4 : Bool;
      _w5 : Bool;
      _w6 : Bool;
      _w7 : Bool;
      _w8 : Bool;
      _w9 : Bool;
      _w10 : Bool;
      _w11 : Bool;
      _w12 : Bool;
      _w13 : Bool;
      _w14 : Bool;
      _w15 : Bool;
   END_VAR
BEGIN

REGION Network 1: START PLC
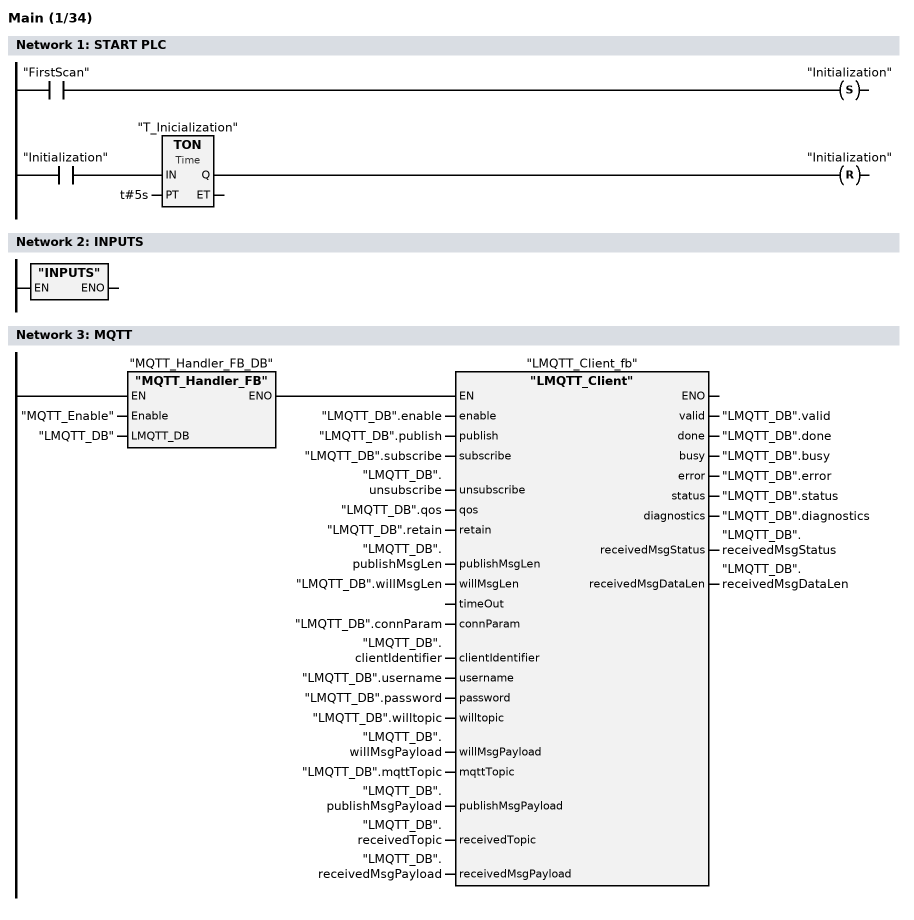
   RUNG wire#powerrail
      Contact( "FirstScan" )
      S_Coil( "Initialization" )
   END_RUNG
   RUNG wire#powerrail
      Contact( "Initialization" )
      { S7_Templates := "time_type := Time" } "T_Inicialization".TON(pt := t#5s, et =>)
      R_Coil( "Initialization" )
   END_RUNG
   // the same network as SCL:
   IF "FirstScan" THEN "Initialization" := TRUE; END_IF;
   "T_Inicialization".TON(IN := "Initialization", PT := t#5s);
   IF "T_Inicialization".Q THEN "Initialization" := FALSE; END_IF;
END_REGION

REGION Network 2: INPUTS
   RUNG wire#powerrail
      "INPUTS"()
   END_RUNG
   // the same network as SCL:
   "INPUTS"();
END_REGION

REGION Network 3: MQTT
   RUNG wire#powerrail
      "MQTT_Handler_FB_DB"(Enable := "MQTT_Enable", LMQTT_DB := "LMQTT_DB")
      "LMQTT_Client_fb"(enable := "LMQTT_DB".enable, publish := "LMQTT_DB".publish, subscribe := "LMQTT_DB".subscribe, unsubscribe := "LMQTT_DB".unsubscribe, qos := "LMQTT_DB".qos, retain := "LMQTT_DB".retain, publishMsgLen := "LMQTT_DB".publishMsgLen, willMsgLen := "LMQTT_DB".willMsgLen, timeOut :=, connParam := "LMQTT_DB".connParam, clientIdentifier := "LMQTT_DB".clientIdentifier, username := "LMQTT_DB".username, password := "LMQTT_DB".password, willtopic := "LMQTT_DB".willtopic, willMsgPayload := "LMQTT_DB".willMsgPayload, mqttTopic := "LMQTT_DB".mqttTopic, publishMsgPayload := "LMQTT_DB".publishMsgPayload, receivedTopic := "LMQTT_DB".receivedTopic, receivedMsgPayload := "LMQTT_DB".receivedMsgPayload, valid => "LMQTT_DB".valid, done => "LMQTT_DB".done, busy => "LMQTT_DB".busy, error => "LMQTT_DB".error, status => "LMQTT_DB".status, diagnostics => "LMQTT_DB".diagnostics, receivedMsgStatus => "LMQTT_DB".receivedMsgStatus, receivedMsgDataLen => "LMQTT_DB".receivedMsgDataLen)
   END_RUNG
   // the same network as SCL:
   "MQTT_Handler_FB_DB"(Enable := "MQTT_Enable", LMQTT_DB := "LMQTT_DB", ENO => #_w1);   // "MQTT_Handler_FB"
   IF #_w1 THEN
       "LMQTT_Client_fb"(enable := "LMQTT_DB".enable,   // "LMQTT_Client"
                         publish := "LMQTT_DB".publish,
                         subscribe := "LMQTT_DB".subscribe,
                         unsubscribe := "LMQTT_DB".unsubscribe,
                         qos := "LMQTT_DB".qos,
                         retain := "LMQTT_DB".retain,
                         publishMsgLen := "LMQTT_DB".publishMsgLen,
                         willMsgLen := "LMQTT_DB".willMsgLen,
                         connParam := "LMQTT_DB".connParam,
                         clientIdentifier := "LMQTT_DB".clientIdentifier,
                         username := "LMQTT_DB".username,
                         password := "LMQTT_DB".password,
                         willtopic := "LMQTT_DB".willtopic,
                         willMsgPayload := "LMQTT_DB".willMsgPayload,
                         mqttTopic := "LMQTT_DB".mqttTopic,
                         publishMsgPayload := "LMQTT_DB".publishMsgPayload,
                         receivedTopic := "LMQTT_DB".receivedTopic,
                         receivedMsgPayload := "LMQTT_DB".receivedMsgPayload,
                         valid => "LMQTT_DB".valid,
                         done => "LMQTT_DB".done,
                         busy => "LMQTT_DB".busy,
                         error => "LMQTT_DB".error,
                         status => "LMQTT_DB".status,
                         diagnostics => "LMQTT_DB".diagnostics,
                         receivedMsgStatus => "LMQTT_DB".receivedMsgStatus,
                         receivedMsgDataLen => "LMQTT_DB".receivedMsgDataLen);
   END_IF;
END_REGION

REGION Network 4: Absolute Encoders
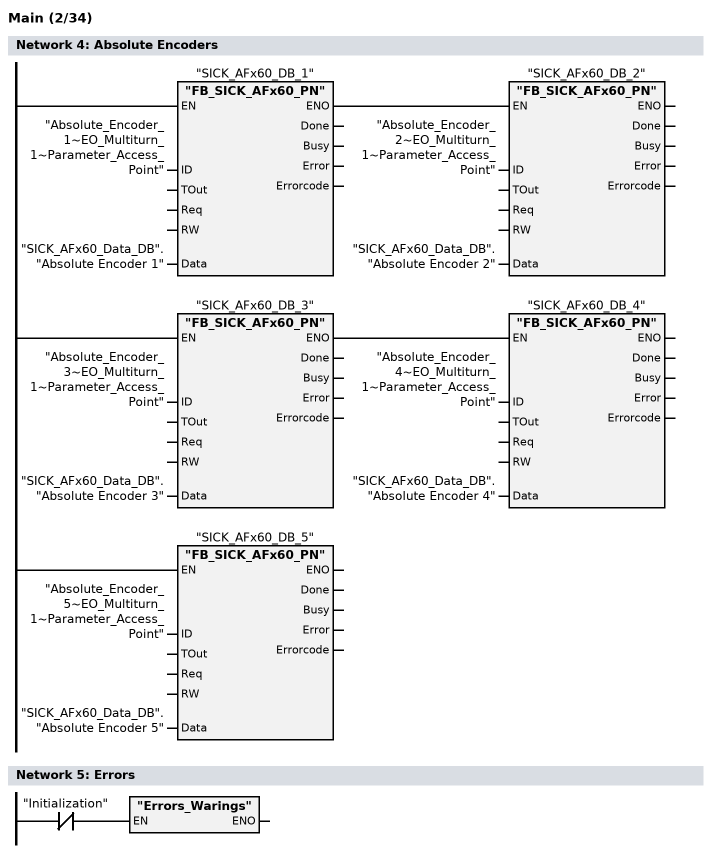
   RUNG wire#powerrail
      "SICK_AFx60_DB_1"(ID := "Absolute_Encoder_1~EO_Multiturn_1~Parameter_Access_Point", TOut :=, Req :=, RW :=, Data := "SICK_AFx60_Data_DB"."Absolute Encoder 1", Done =>, Busy =>, Error =>, Errorcode =>)
      "SICK_AFx60_DB_2"(ID := "Absolute_Encoder_2~EO_Multiturn_1~Parameter_Access_Point", TOut :=, Req :=, RW :=, Data := "SICK_AFx60_Data_DB"."Absolute Encoder 2", Done =>, Busy =>, Error =>, Errorcode =>)
   END_RUNG
   RUNG wire#powerrail
      "SICK_AFx60_DB_3"(ID := "Absolute_Encoder_3~EO_Multiturn_1~Parameter_Access_Point", TOut :=, Req :=, RW :=, Data := "SICK_AFx60_Data_DB"."Absolute Encoder 3", Done =>, Busy =>, Error =>, Errorcode =>)
      "SICK_AFx60_DB_4"(ID := "Absolute_Encoder_4~EO_Multiturn_1~Parameter_Access_Point", TOut :=, Req :=, RW :=, Data := "SICK_AFx60_Data_DB"."Absolute Encoder 4", Done =>, Busy =>, Error =>, Errorcode =>)
   END_RUNG
   RUNG wire#powerrail
      "SICK_AFx60_DB_5"(ID := "Absolute_Encoder_5~EO_Multiturn_1~Parameter_Access_Point", TOut :=, Req :=, RW :=, Data := "SICK_AFx60_Data_DB"."Absolute Encoder 5", Done =>, Busy =>, Error =>, Errorcode =>)
   END_RUNG
   // the same network as SCL:
   "SICK_AFx60_DB_1"(ID := "Absolute_Encoder_1~EO_Multiturn_1~Parameter_Access_Point",   // "FB_SICK_AFx60_PN"
                     Data := "SICK_AFx60_Data_DB"."Absolute Encoder 1",
                     ENO => #_w1);
   IF #_w1 THEN
       "SICK_AFx60_DB_2"(ID := "Absolute_Encoder_2~EO_Multiturn_1~Parameter_Access_Point",   // "FB_SICK_AFx60_PN"
                         Data := "SICK_AFx60_Data_DB"."Absolute Encoder 2");
   END_IF;
   "SICK_AFx60_DB_3"(ID := "Absolute_Encoder_3~EO_Multiturn_1~Parameter_Access_Point",   // "FB_SICK_AFx60_PN"
                     Data := "SICK_AFx60_Data_DB"."Absolute Encoder 3",
                     ENO => #_w2);
   IF #_w2 THEN
       "SICK_AFx60_DB_4"(ID := "Absolute_Encoder_4~EO_Multiturn_1~Parameter_Access_Point",   // "FB_SICK_AFx60_PN"
                         Data := "SICK_AFx60_Data_DB"."Absolute Encoder 4");
   END_IF;
   "SICK_AFx60_DB_5"(ID := "Absolute_Encoder_5~EO_Multiturn_1~Parameter_Access_Point",   // "FB_SICK_AFx60_PN"
                     Data := "SICK_AFx60_Data_DB"."Absolute Encoder 5");
END_REGION

REGION Network 5: Errors
   RUNG wire#powerrail
      I_Contact( "Initialization" )
      "Errors_Warings"()
   END_RUNG
   // the same network as SCL:
   IF NOT "Initialization" THEN "Errors_Warings"(); END_IF;
END_REGION

REGION Network 6: AUTO TEST 1
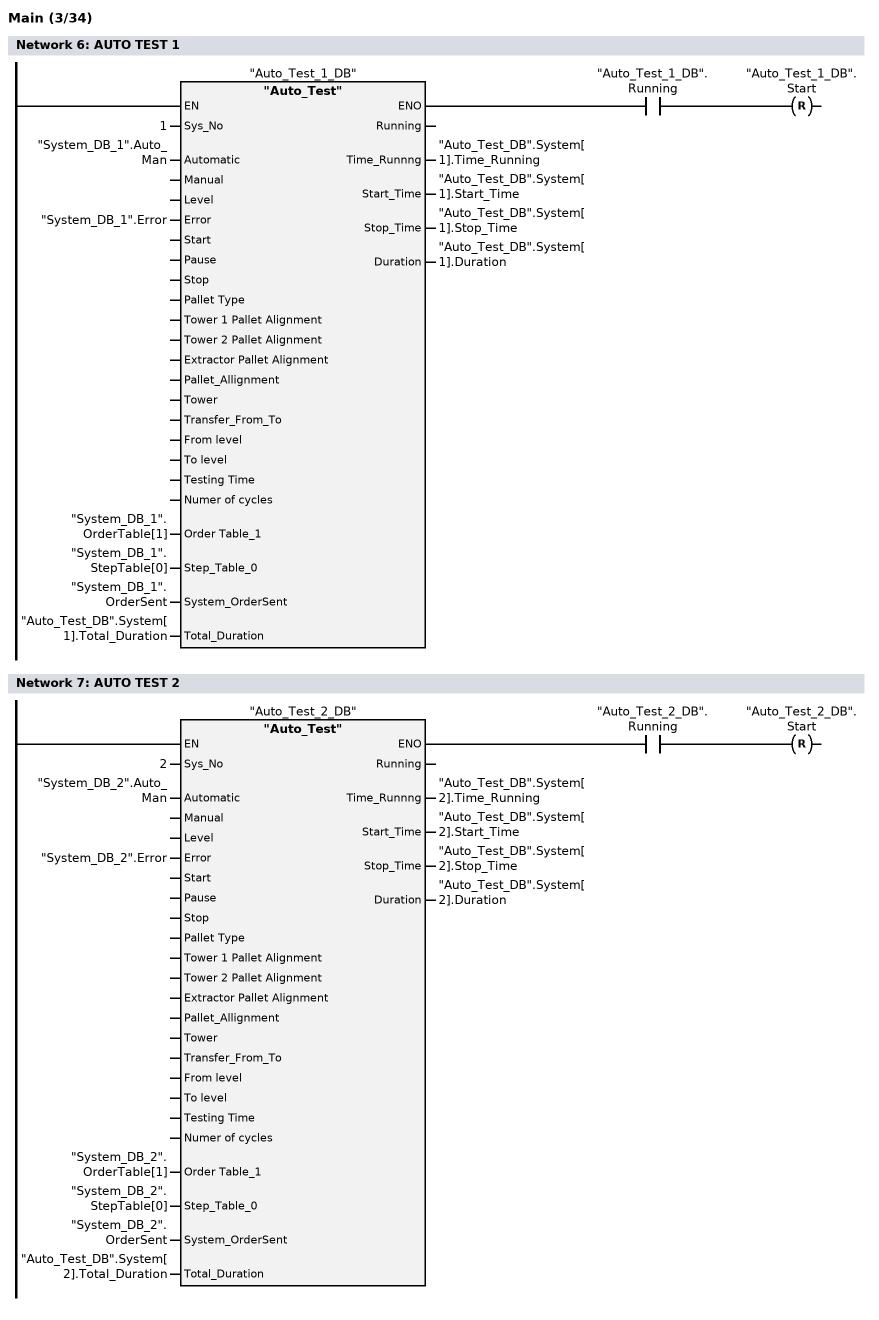
   RUNG wire#powerrail
      "Auto_Test_1_DB"(Sys_No := 1, Automatic := "System_DB_1".Auto_Man, Manual :=, Level :=, Error := "System_DB_1".Error, Start :=, Pause :=, Stop :=, "Pallet Type" :=, "Tower 1 Pallet Alignment" :=, "Tower 2 Pallet Alignment" :=, "Extractor Pallet Alignment" :=, Pallet_Allignment :=, Tower :=, Transfer_From_To :=, "From level" :=, "To level" :=, "Testing Time" :=, "Numer of cycles" :=, "Order Table_1" := "System_DB_1".OrderTable[1], Step_Table_0 := "System_DB_1".StepTable[0], System_OrderSent := "System_DB_1".OrderSent, Total_Duration := "Auto_Test_DB".System[1].Total_Duration, Running =>, Time_Runnng => "Auto_Test_DB".System[1].Time_Running, Start_Time => "Auto_Test_DB".System[1].Start_Time, Stop_Time => "Auto_Test_DB".System[1].Stop_Time, Duration => "Auto_Test_DB".System[1].Duration)
      Contact( "Auto_Test_1_DB".Running )
      R_Coil( "Auto_Test_1_DB".Start )
   END_RUNG
   // the same network as SCL:
   "Auto_Test_1_DB"(Sys_No := 1,   // "Auto_Test"
                    Automatic := "System_DB_1".Auto_Man,
                    Error := "System_DB_1".Error,
                    "Order Table_1" := "System_DB_1".OrderTable[1],
                    Step_Table_0 := "System_DB_1".StepTable[0],
                    System_OrderSent := "System_DB_1".OrderSent,
                    Total_Duration := "Auto_Test_DB".System[1].Total_Duration,
                    Time_Runnng => "Auto_Test_DB".System[1].Time_Running,
                    Start_Time => "Auto_Test_DB".System[1].Start_Time,
                    Stop_Time => "Auto_Test_DB".System[1].Stop_Time,
                    Duration => "Auto_Test_DB".System[1].Duration,
                    ENO => #_w1);
   IF #_w1 AND "Auto_Test_1_DB".Running THEN "Auto_Test_1_DB".Start := FALSE; END_IF;
END_REGION

REGION Network 7: AUTO TEST 2
   RUNG wire#powerrail
      "Auto_Test_2_DB"(Sys_No := 2, Automatic := "System_DB_2".Auto_Man, Manual :=, Level :=, Error := "System_DB_2".Error, Start :=, Pause :=, Stop :=, "Pallet Type" :=, "Tower 1 Pallet Alignment" :=, "Tower 2 Pallet Alignment" :=, "Extractor Pallet Alignment" :=, Pallet_Allignment :=, Tower :=, Transfer_From_To :=, "From level" :=, "To level" :=, "Testing Time" :=, "Numer of cycles" :=, "Order Table_1" := "System_DB_2".OrderTable[1], Step_Table_0 := "System_DB_2".StepTable[0], System_OrderSent := "System_DB_2".OrderSent, Total_Duration := "Auto_Test_DB".System[2].Total_Duration, Running =>, Time_Runnng => "Auto_Test_DB".System[2].Time_Running, Start_Time => "Auto_Test_DB".System[2].Start_Time, Stop_Time => "Auto_Test_DB".System[2].Stop_Time, Duration => "Auto_Test_DB".System[2].Duration)
      Contact( "Auto_Test_2_DB".Running )
      R_Coil( "Auto_Test_2_DB".Start )
   END_RUNG
   // the same network as SCL:
   "Auto_Test_2_DB"(Sys_No := 2,   // "Auto_Test"
                    Automatic := "System_DB_2".Auto_Man,
                    Error := "System_DB_2".Error,
                    "Order Table_1" := "System_DB_2".OrderTable[1],
                    Step_Table_0 := "System_DB_2".StepTable[0],
                    System_OrderSent := "System_DB_2".OrderSent,
                    Total_Duration := "Auto_Test_DB".System[2].Total_Duration,
                    Time_Runnng => "Auto_Test_DB".System[2].Time_Running,
                    Start_Time => "Auto_Test_DB".System[2].Start_Time,
                    Stop_Time => "Auto_Test_DB".System[2].Stop_Time,
                    Duration => "Auto_Test_DB".System[2].Duration,
                    ENO => #_w1);
   IF #_w1 AND "Auto_Test_2_DB".Running THEN "Auto_Test_2_DB".Start := FALSE; END_IF;
END_REGION

REGION Network 8: AUTO TEST 3
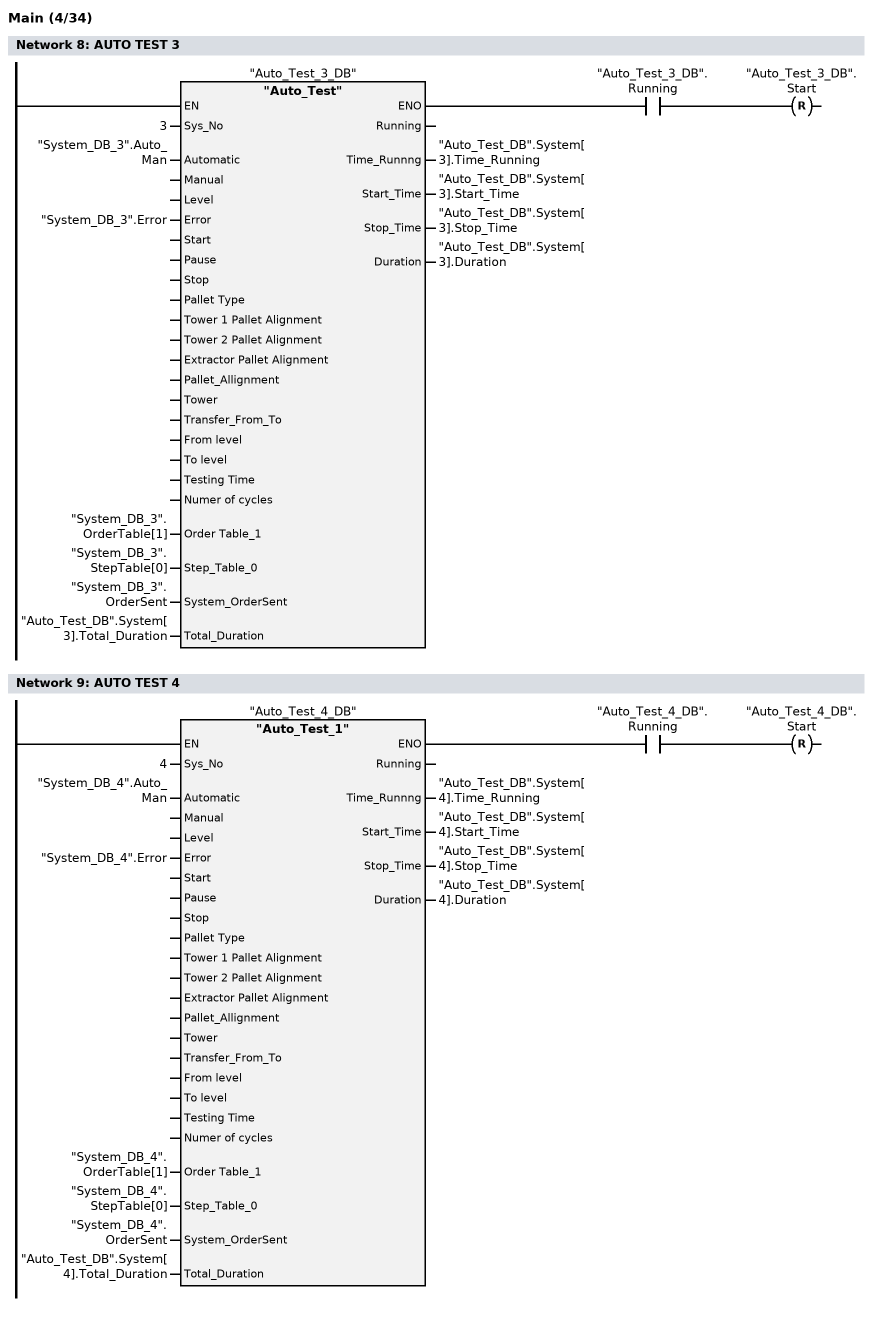
   RUNG wire#powerrail
      "Auto_Test_3_DB"(Sys_No := 3, Automatic := "System_DB_3".Auto_Man, Manual :=, Level :=, Error := "System_DB_3".Error, Start :=, Pause :=, Stop :=, "Pallet Type" :=, "Tower 1 Pallet Alignment" :=, "Tower 2 Pallet Alignment" :=, "Extractor Pallet Alignment" :=, Pallet_Allignment :=, Tower :=, Transfer_From_To :=, "From level" :=, "To level" :=, "Testing Time" :=, "Numer of cycles" :=, "Order Table_1" := "System_DB_3".OrderTable[1], Step_Table_0 := "System_DB_3".StepTable[0], System_OrderSent := "System_DB_3".OrderSent, Total_Duration := "Auto_Test_DB".System[3].Total_Duration, Running =>, Time_Runnng => "Auto_Test_DB".System[3].Time_Running, Start_Time => "Auto_Test_DB".System[3].Start_Time, Stop_Time => "Auto_Test_DB".System[3].Stop_Time, Duration => "Auto_Test_DB".System[3].Duration)
      Contact( "Auto_Test_3_DB".Running )
      R_Coil( "Auto_Test_3_DB".Start )
   END_RUNG
   // the same network as SCL:
   "Auto_Test_3_DB"(Sys_No := 3,   // "Auto_Test"
                    Automatic := "System_DB_3".Auto_Man,
                    Error := "System_DB_3".Error,
                    "Order Table_1" := "System_DB_3".OrderTable[1],
                    Step_Table_0 := "System_DB_3".StepTable[0],
                    System_OrderSent := "System_DB_3".OrderSent,
                    Total_Duration := "Auto_Test_DB".System[3].Total_Duration,
                    Time_Runnng => "Auto_Test_DB".System[3].Time_Running,
                    Start_Time => "Auto_Test_DB".System[3].Start_Time,
                    Stop_Time => "Auto_Test_DB".System[3].Stop_Time,
                    Duration => "Auto_Test_DB".System[3].Duration,
                    ENO => #_w1);
   IF #_w1 AND "Auto_Test_3_DB".Running THEN "Auto_Test_3_DB".Start := FALSE; END_IF;
END_REGION

REGION Network 9: AUTO TEST 4
   RUNG wire#powerrail
      "Auto_Test_4_DB"(Sys_No := 4, Automatic := "System_DB_4".Auto_Man, Manual :=, Level :=, Error := "System_DB_4".Error, Start :=, Pause :=, Stop :=, "Pallet Type" :=, "Tower 1 Pallet Alignment" :=, "Tower 2 Pallet Alignment" :=, "Extractor Pallet Alignment" :=, Pallet_Allignment :=, Tower :=, Transfer_From_To :=, "From level" :=, "To level" :=, "Testing Time" :=, "Numer of cycles" :=, "Order Table_1" := "System_DB_4".OrderTable[1], Step_Table_0 := "System_DB_4".StepTable[0], System_OrderSent := "System_DB_4".OrderSent, Total_Duration := "Auto_Test_DB".System[4].Total_Duration, Running =>, Time_Runnng => "Auto_Test_DB".System[4].Time_Running, Start_Time => "Auto_Test_DB".System[4].Start_Time, Stop_Time => "Auto_Test_DB".System[4].Stop_Time, Duration => "Auto_Test_DB".System[4].Duration)
      Contact( "Auto_Test_4_DB".Running )
      R_Coil( "Auto_Test_4_DB".Start )
   END_RUNG
   // the same network as SCL:
   "Auto_Test_4_DB"(Sys_No := 4,   // "Auto_Test_1"
                    Automatic := "System_DB_4".Auto_Man,
                    Error := "System_DB_4".Error,
                    "Order Table_1" := "System_DB_4".OrderTable[1],
                    Step_Table_0 := "System_DB_4".StepTable[0],
                    System_OrderSent := "System_DB_4".OrderSent,
                    Total_Duration := "Auto_Test_DB".System[4].Total_Duration,
                    Time_Runnng => "Auto_Test_DB".System[4].Time_Running,
                    Start_Time => "Auto_Test_DB".System[4].Start_Time,
                    Stop_Time => "Auto_Test_DB".System[4].Stop_Time,
                    Duration => "Auto_Test_DB".System[4].Duration,
                    ENO => #_w1);
   IF #_w1 AND "Auto_Test_4_DB".Running THEN "Auto_Test_4_DB".Start := FALSE; END_IF;
END_REGION

REGION Network 10: AUTO TEST 5
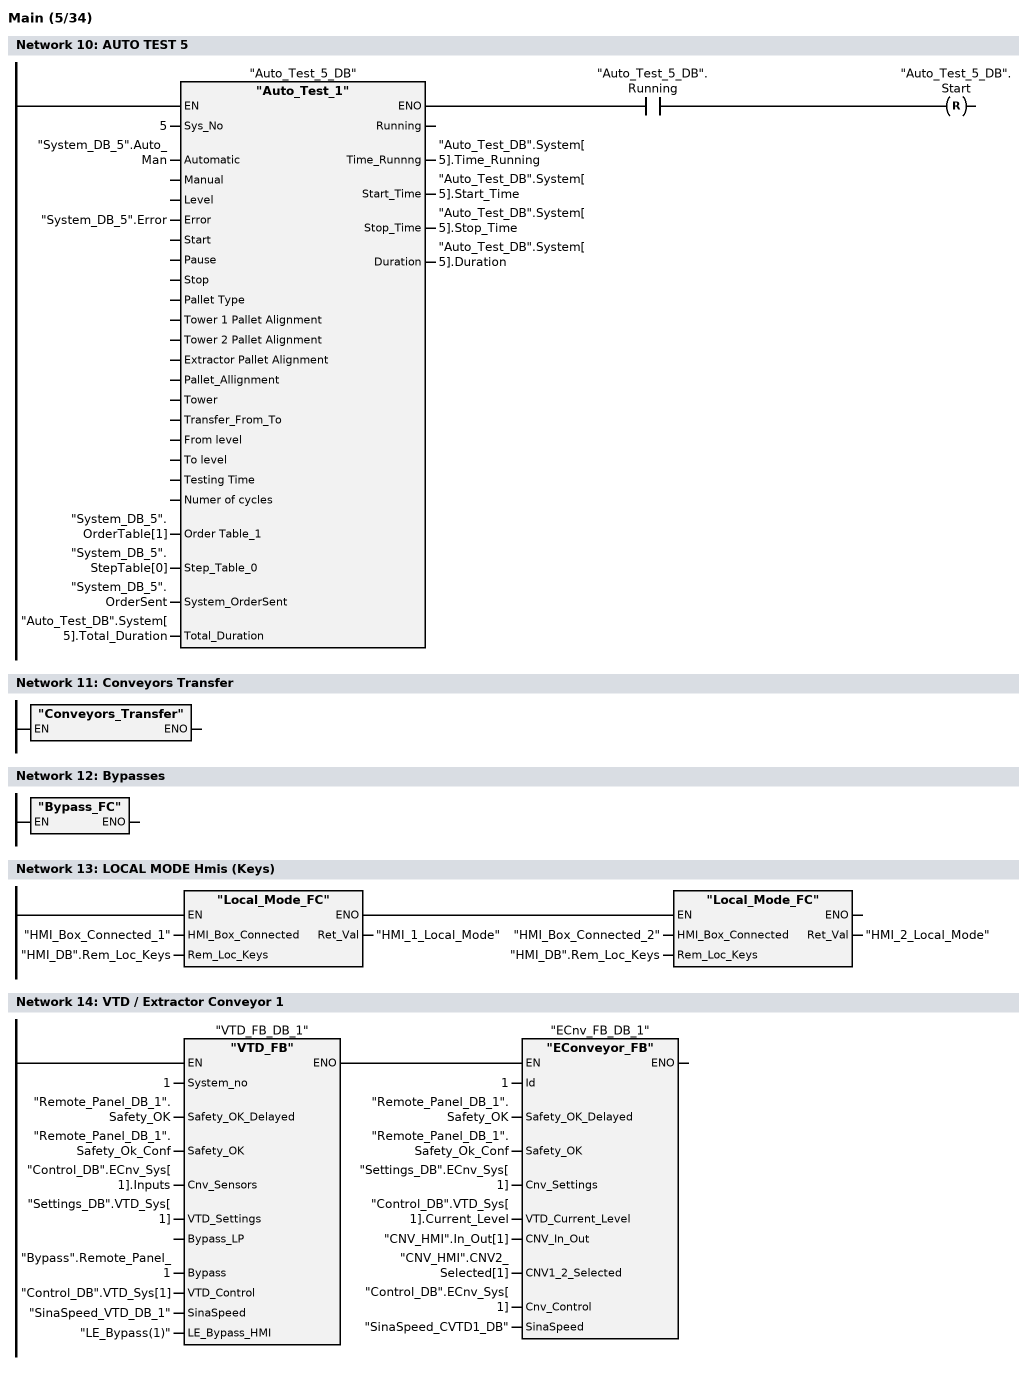
   RUNG wire#powerrail
      "Auto_Test_5_DB"(Sys_No := 5, Automatic := "System_DB_5".Auto_Man, Manual :=, Level :=, Error := "System_DB_5".Error, Start :=, Pause :=, Stop :=, "Pallet Type" :=, "Tower 1 Pallet Alignment" :=, "Tower 2 Pallet Alignment" :=, "Extractor Pallet Alignment" :=, Pallet_Allignment :=, Tower :=, Transfer_From_To :=, "From level" :=, "To level" :=, "Testing Time" :=, "Numer of cycles" :=, "Order Table_1" := "System_DB_5".OrderTable[1], Step_Table_0 := "System_DB_5".StepTable[0], System_OrderSent := "System_DB_5".OrderSent, Total_Duration := "Auto_Test_DB".System[5].Total_Duration, Running =>, Time_Runnng => "Auto_Test_DB".System[5].Time_Running, Start_Time => "Auto_Test_DB".System[5].Start_Time, Stop_Time => "Auto_Test_DB".System[5].Stop_Time, Duration => "Auto_Test_DB".System[5].Duration)
      Contact( "Auto_Test_5_DB".Running )
      R_Coil( "Auto_Test_5_DB".Start )
   END_RUNG
   // the same network as SCL:
   "Auto_Test_5_DB"(Sys_No := 5,   // "Auto_Test_1"
                    Automatic := "System_DB_5".Auto_Man,
                    Error := "System_DB_5".Error,
                    "Order Table_1" := "System_DB_5".OrderTable[1],
                    Step_Table_0 := "System_DB_5".StepTable[0],
                    System_OrderSent := "System_DB_5".OrderSent,
                    Total_Duration := "Auto_Test_DB".System[5].Total_Duration,
                    Time_Runnng => "Auto_Test_DB".System[5].Time_Running,
                    Start_Time => "Auto_Test_DB".System[5].Start_Time,
                    Stop_Time => "Auto_Test_DB".System[5].Stop_Time,
                    Duration => "Auto_Test_DB".System[5].Duration,
                    ENO => #_w1);
   IF #_w1 AND "Auto_Test_5_DB".Running THEN "Auto_Test_5_DB".Start := FALSE; END_IF;
END_REGION

REGION Network 11: Conveyors Transfer
   RUNG wire#powerrail
      "Conveyors_Transfer"()
   END_RUNG
   // the same network as SCL:
   "Conveyors_Transfer"();
END_REGION

REGION Network 12: Bypasses
   RUNG wire#powerrail
      "Bypass_FC"()
   END_RUNG
   // the same network as SCL:
   "Bypass_FC"();
END_REGION

REGION Network 13: LOCAL MODE Hmis (Keys)
   RUNG wire#powerrail
      "Local_Mode_FC"(HMI_Box_Connected := "HMI_Box_Connected_1", Rem_Loc_Keys := "HMI_DB".Rem_Loc_Keys, Ret_Val => "HMI_1_Local_Mode")
      "Local_Mode_FC"(HMI_Box_Connected := "HMI_Box_Connected_2", Rem_Loc_Keys := "HMI_DB".Rem_Loc_Keys, Ret_Val => "HMI_2_Local_Mode")
   END_RUNG
   // the same network as SCL:
   "HMI_1_Local_Mode" := "Local_Mode_FC"(HMI_Box_Connected := "HMI_Box_Connected_1",
                           Rem_Loc_Keys := "HMI_DB".Rem_Loc_Keys,
                           ENO => #_w1);
   IF #_w1 THEN
       "HMI_2_Local_Mode" := "Local_Mode_FC"(HMI_Box_Connected := "HMI_Box_Connected_2",
                               Rem_Loc_Keys := "HMI_DB".Rem_Loc_Keys);
   END_IF;
END_REGION

REGION Network 14: VTD / Extractor Conveyor 1
   RUNG wire#powerrail
      "VTD_FB_DB_1"(System_no := 1, Safety_OK_Delayed := "Remote_Panel_DB_1".Safety_OK, Safety_OK := "Remote_Panel_DB_1".Safety_Ok_Conf, Cnv_Sensors := "Control_DB".ECnv_Sys[1].Inputs, VTD_Settings := "Settings_DB".VTD_Sys[1], Bypass_LP :=, Bypass := "Bypass".Remote_Panel_1, VTD_Control := "Control_DB".VTD_Sys[1], SinaSpeed := "SinaSpeed_VTD_DB_1", LE_Bypass_HMI := "LE_Bypass(1)")
      "ECnv_FB_DB_1"(Id := 1, Safety_OK_Delayed := "Remote_Panel_DB_1".Safety_OK, Safety_OK := "Remote_Panel_DB_1".Safety_Ok_Conf, Cnv_Settings := "Settings_DB".ECnv_Sys[1], VTD_Current_Level := "Control_DB".VTD_Sys[1].Current_Level, CNV_In_Out := "CNV_HMI".In_Out[1], CNV1_2_Selected := "CNV_HMI".CNV2_Selected[1], Cnv_Control := "Control_DB".ECnv_Sys[1], SinaSpeed := "SinaSpeed_CVTD1_DB")
   END_RUNG
   // the same network as SCL:
   "VTD_FB_DB_1"(System_no := 1,   // "VTD_FB"
                 Safety_OK_Delayed := "Remote_Panel_DB_1".Safety_OK,
                 Safety_OK := "Remote_Panel_DB_1".Safety_Ok_Conf,
                 Cnv_Sensors := "Control_DB".ECnv_Sys[1].Inputs,
                 VTD_Settings := "Settings_DB".VTD_Sys[1],
                 Bypass := "Bypass".Remote_Panel_1,
                 VTD_Control := "Control_DB".VTD_Sys[1],
                 SinaSpeed := "SinaSpeed_VTD_DB_1",
                 LE_Bypass_HMI := "LE_Bypass(1)",
                 ENO => #_w1);
   IF #_w1 THEN
       "ECnv_FB_DB_1"(Id := 1,   // "EConveyor_FB"
                      Safety_OK_Delayed := "Remote_Panel_DB_1".Safety_OK,
                      Safety_OK := "Remote_Panel_DB_1".Safety_Ok_Conf,
                      Cnv_Settings := "Settings_DB".ECnv_Sys[1],
                      VTD_Current_Level := "Control_DB".VTD_Sys[1].Current_Level,
                      CNV_In_Out := "CNV_HMI".In_Out[1],
                      CNV1_2_Selected := "CNV_HMI".CNV2_Selected[1],
                      Cnv_Control := "Control_DB".ECnv_Sys[1],
                      SinaSpeed := "SinaSpeed_CVTD1_DB");
   END_IF;
END_REGION

REGION Network 15: VTD / Extractor Conveyor 2
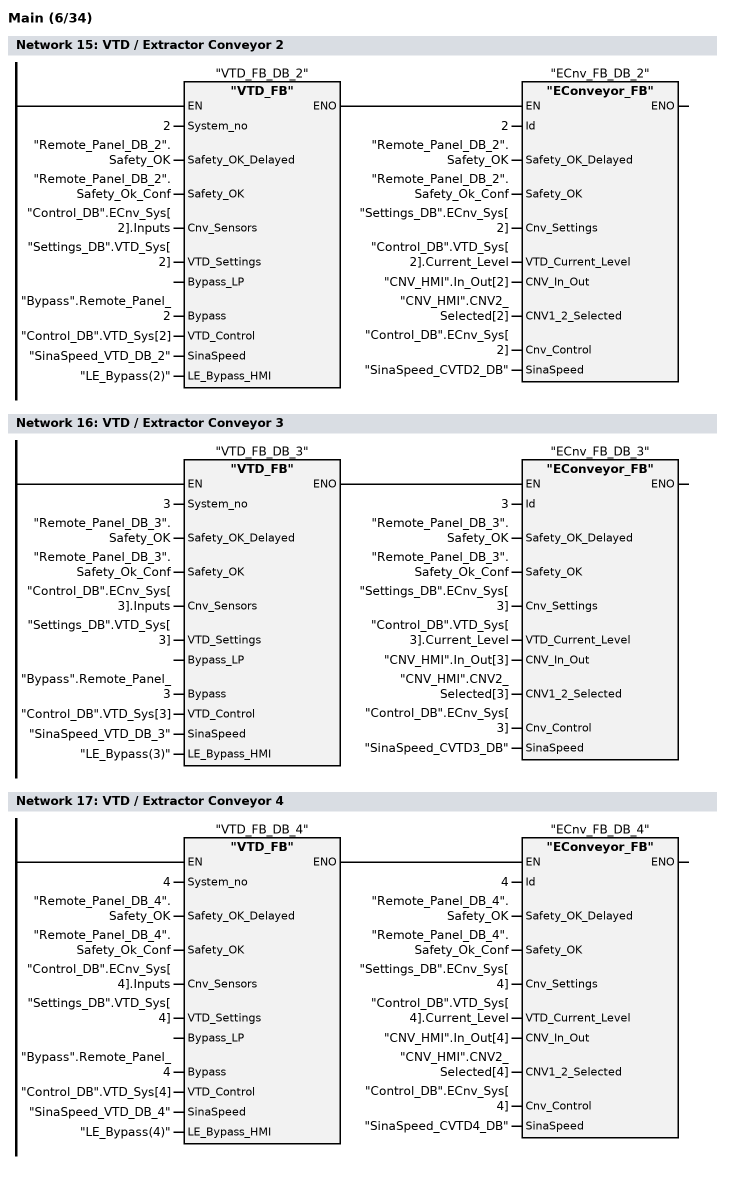
   RUNG wire#powerrail
      "VTD_FB_DB_2"(System_no := 2, Safety_OK_Delayed := "Remote_Panel_DB_2".Safety_OK, Safety_OK := "Remote_Panel_DB_2".Safety_Ok_Conf, Cnv_Sensors := "Control_DB".ECnv_Sys[2].Inputs, VTD_Settings := "Settings_DB".VTD_Sys[2], Bypass_LP :=, Bypass := "Bypass".Remote_Panel_2, VTD_Control := "Control_DB".VTD_Sys[2], SinaSpeed := "SinaSpeed_VTD_DB_2", LE_Bypass_HMI := "LE_Bypass(2)")
      "ECnv_FB_DB_2"(Id := 2, Safety_OK_Delayed := "Remote_Panel_DB_2".Safety_OK, Safety_OK := "Remote_Panel_DB_2".Safety_Ok_Conf, Cnv_Settings := "Settings_DB".ECnv_Sys[2], VTD_Current_Level := "Control_DB".VTD_Sys[2].Current_Level, CNV_In_Out := "CNV_HMI".In_Out[2], CNV1_2_Selected := "CNV_HMI".CNV2_Selected[2], Cnv_Control := "Control_DB".ECnv_Sys[2], SinaSpeed := "SinaSpeed_CVTD2_DB")
   END_RUNG
   // the same network as SCL:
   "VTD_FB_DB_2"(System_no := 2,   // "VTD_FB"
                 Safety_OK_Delayed := "Remote_Panel_DB_2".Safety_OK,
                 Safety_OK := "Remote_Panel_DB_2".Safety_Ok_Conf,
                 Cnv_Sensors := "Control_DB".ECnv_Sys[2].Inputs,
                 VTD_Settings := "Settings_DB".VTD_Sys[2],
                 Bypass := "Bypass".Remote_Panel_2,
                 VTD_Control := "Control_DB".VTD_Sys[2],
                 SinaSpeed := "SinaSpeed_VTD_DB_2",
                 LE_Bypass_HMI := "LE_Bypass(2)",
                 ENO => #_w1);
   IF #_w1 THEN
       "ECnv_FB_DB_2"(Id := 2,   // "EConveyor_FB"
                      Safety_OK_Delayed := "Remote_Panel_DB_2".Safety_OK,
                      Safety_OK := "Remote_Panel_DB_2".Safety_Ok_Conf,
                      Cnv_Settings := "Settings_DB".ECnv_Sys[2],
                      VTD_Current_Level := "Control_DB".VTD_Sys[2].Current_Level,
                      CNV_In_Out := "CNV_HMI".In_Out[2],
                      CNV1_2_Selected := "CNV_HMI".CNV2_Selected[2],
                      Cnv_Control := "Control_DB".ECnv_Sys[2],
                      SinaSpeed := "SinaSpeed_CVTD2_DB");
   END_IF;
END_REGION

REGION Network 16: VTD / Extractor Conveyor 3
   RUNG wire#powerrail
      "VTD_FB_DB_3"(System_no := 3, Safety_OK_Delayed := "Remote_Panel_DB_3".Safety_OK, Safety_OK := "Remote_Panel_DB_3".Safety_Ok_Conf, Cnv_Sensors := "Control_DB".ECnv_Sys[3].Inputs, VTD_Settings := "Settings_DB".VTD_Sys[3], Bypass_LP :=, Bypass := "Bypass".Remote_Panel_3, VTD_Control := "Control_DB".VTD_Sys[3], SinaSpeed := "SinaSpeed_VTD_DB_3", LE_Bypass_HMI := "LE_Bypass(3)")
      "ECnv_FB_DB_3"(Id := 3, Safety_OK_Delayed := "Remote_Panel_DB_3".Safety_OK, Safety_OK := "Remote_Panel_DB_3".Safety_Ok_Conf, Cnv_Settings := "Settings_DB".ECnv_Sys[3], VTD_Current_Level := "Control_DB".VTD_Sys[3].Current_Level, CNV_In_Out := "CNV_HMI".In_Out[3], CNV1_2_Selected := "CNV_HMI".CNV2_Selected[3], Cnv_Control := "Control_DB".ECnv_Sys[3], SinaSpeed := "SinaSpeed_CVTD3_DB")
   END_RUNG
   // the same network as SCL:
   "VTD_FB_DB_3"(System_no := 3,   // "VTD_FB"
                 Safety_OK_Delayed := "Remote_Panel_DB_3".Safety_OK,
                 Safety_OK := "Remote_Panel_DB_3".Safety_Ok_Conf,
                 Cnv_Sensors := "Control_DB".ECnv_Sys[3].Inputs,
                 VTD_Settings := "Settings_DB".VTD_Sys[3],
                 Bypass := "Bypass".Remote_Panel_3,
                 VTD_Control := "Control_DB".VTD_Sys[3],
                 SinaSpeed := "SinaSpeed_VTD_DB_3",
                 LE_Bypass_HMI := "LE_Bypass(3)",
                 ENO => #_w1);
   IF #_w1 THEN
       "ECnv_FB_DB_3"(Id := 3,   // "EConveyor_FB"
                      Safety_OK_Delayed := "Remote_Panel_DB_3".Safety_OK,
                      Safety_OK := "Remote_Panel_DB_3".Safety_Ok_Conf,
                      Cnv_Settings := "Settings_DB".ECnv_Sys[3],
                      VTD_Current_Level := "Control_DB".VTD_Sys[3].Current_Level,
                      CNV_In_Out := "CNV_HMI".In_Out[3],
                      CNV1_2_Selected := "CNV_HMI".CNV2_Selected[3],
                      Cnv_Control := "Control_DB".ECnv_Sys[3],
                      SinaSpeed := "SinaSpeed_CVTD3_DB");
   END_IF;
END_REGION

REGION Network 17: VTD / Extractor Conveyor 4
   RUNG wire#powerrail
      "VTD_FB_DB_4"(System_no := 4, Safety_OK_Delayed := "Remote_Panel_DB_4".Safety_OK, Safety_OK := "Remote_Panel_DB_4".Safety_Ok_Conf, Cnv_Sensors := "Control_DB".ECnv_Sys[4].Inputs, VTD_Settings := "Settings_DB".VTD_Sys[4], Bypass_LP :=, Bypass := "Bypass".Remote_Panel_4, VTD_Control := "Control_DB".VTD_Sys[4], SinaSpeed := "SinaSpeed_VTD_DB_4", LE_Bypass_HMI := "LE_Bypass(4)")
      "ECnv_FB_DB_4"(Id := 4, Safety_OK_Delayed := "Remote_Panel_DB_4".Safety_OK, Safety_OK := "Remote_Panel_DB_4".Safety_Ok_Conf, Cnv_Settings := "Settings_DB".ECnv_Sys[4], VTD_Current_Level := "Control_DB".VTD_Sys[4].Current_Level, CNV_In_Out := "CNV_HMI".In_Out[4], CNV1_2_Selected := "CNV_HMI".CNV2_Selected[4], Cnv_Control := "Control_DB".ECnv_Sys[4], SinaSpeed := "SinaSpeed_CVTD4_DB")
   END_RUNG
   // the same network as SCL:
   "VTD_FB_DB_4"(System_no := 4,   // "VTD_FB"
                 Safety_OK_Delayed := "Remote_Panel_DB_4".Safety_OK,
                 Safety_OK := "Remote_Panel_DB_4".Safety_Ok_Conf,
                 Cnv_Sensors := "Control_DB".ECnv_Sys[4].Inputs,
                 VTD_Settings := "Settings_DB".VTD_Sys[4],
                 Bypass := "Bypass".Remote_Panel_4,
                 VTD_Control := "Control_DB".VTD_Sys[4],
                 SinaSpeed := "SinaSpeed_VTD_DB_4",
                 LE_Bypass_HMI := "LE_Bypass(4)",
                 ENO => #_w1);
   IF #_w1 THEN
       "ECnv_FB_DB_4"(Id := 4,   // "EConveyor_FB"
                      Safety_OK_Delayed := "Remote_Panel_DB_4".Safety_OK,
                      Safety_OK := "Remote_Panel_DB_4".Safety_Ok_Conf,
                      Cnv_Settings := "Settings_DB".ECnv_Sys[4],
                      VTD_Current_Level := "Control_DB".VTD_Sys[4].Current_Level,
                      CNV_In_Out := "CNV_HMI".In_Out[4],
                      CNV1_2_Selected := "CNV_HMI".CNV2_Selected[4],
                      Cnv_Control := "Control_DB".ECnv_Sys[4],
                      SinaSpeed := "SinaSpeed_CVTD4_DB");
   END_IF;
END_REGION

REGION Network 18: VTD / Extractor Conveyor 5
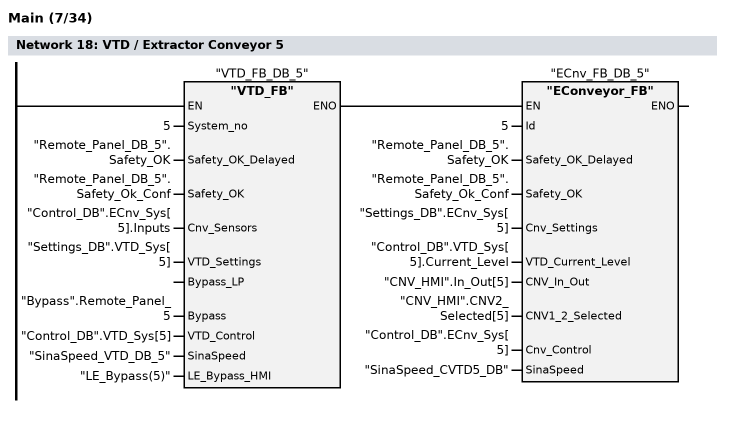
   RUNG wire#powerrail
      "VTD_FB_DB_5"(System_no := 5, Safety_OK_Delayed := "Remote_Panel_DB_5".Safety_OK, Safety_OK := "Remote_Panel_DB_5".Safety_Ok_Conf, Cnv_Sensors := "Control_DB".ECnv_Sys[5].Inputs, VTD_Settings := "Settings_DB".VTD_Sys[5], Bypass_LP :=, Bypass := "Bypass".Remote_Panel_5, VTD_Control := "Control_DB".VTD_Sys[5], SinaSpeed := "SinaSpeed_VTD_DB_5", LE_Bypass_HMI := "LE_Bypass(5)")
      "ECnv_FB_DB_5"(Id := 5, Safety_OK_Delayed := "Remote_Panel_DB_5".Safety_OK, Safety_OK := "Remote_Panel_DB_5".Safety_Ok_Conf, Cnv_Settings := "Settings_DB".ECnv_Sys[5], VTD_Current_Level := "Control_DB".VTD_Sys[5].Current_Level, CNV_In_Out := "CNV_HMI".In_Out[5], CNV1_2_Selected := "CNV_HMI".CNV2_Selected[5], Cnv_Control := "Control_DB".ECnv_Sys[5], SinaSpeed := "SinaSpeed_CVTD5_DB")
   END_RUNG
   // the same network as SCL:
   "VTD_FB_DB_5"(System_no := 5,   // "VTD_FB"
                 Safety_OK_Delayed := "Remote_Panel_DB_5".Safety_OK,
                 Safety_OK := "Remote_Panel_DB_5".Safety_Ok_Conf,
                 Cnv_Sensors := "Control_DB".ECnv_Sys[5].Inputs,
                 VTD_Settings := "Settings_DB".VTD_Sys[5],
                 Bypass := "Bypass".Remote_Panel_5,
                 VTD_Control := "Control_DB".VTD_Sys[5],
                 SinaSpeed := "SinaSpeed_VTD_DB_5",
                 LE_Bypass_HMI := "LE_Bypass(5)",
                 ENO => #_w1);
   IF #_w1 THEN
       "ECnv_FB_DB_5"(Id := 5,   // "EConveyor_FB"
                      Safety_OK_Delayed := "Remote_Panel_DB_5".Safety_OK,
                      Safety_OK := "Remote_Panel_DB_5".Safety_Ok_Conf,
                      Cnv_Settings := "Settings_DB".ECnv_Sys[5],
                      VTD_Current_Level := "Control_DB".VTD_Sys[5].Current_Level,
                      CNV_In_Out := "CNV_HMI".In_Out[5],
                      CNV1_2_Selected := "CNV_HMI".CNV2_Selected[5],
                      Cnv_Control := "Control_DB".ECnv_Sys[5],
                      SinaSpeed := "SinaSpeed_CVTD5_DB");
   END_IF;
END_REGION

REGION Network 19: SYSTEM 1
END_REGION

REGION Network 20: Level Conveyors Tower 1 - SYSTEM 1
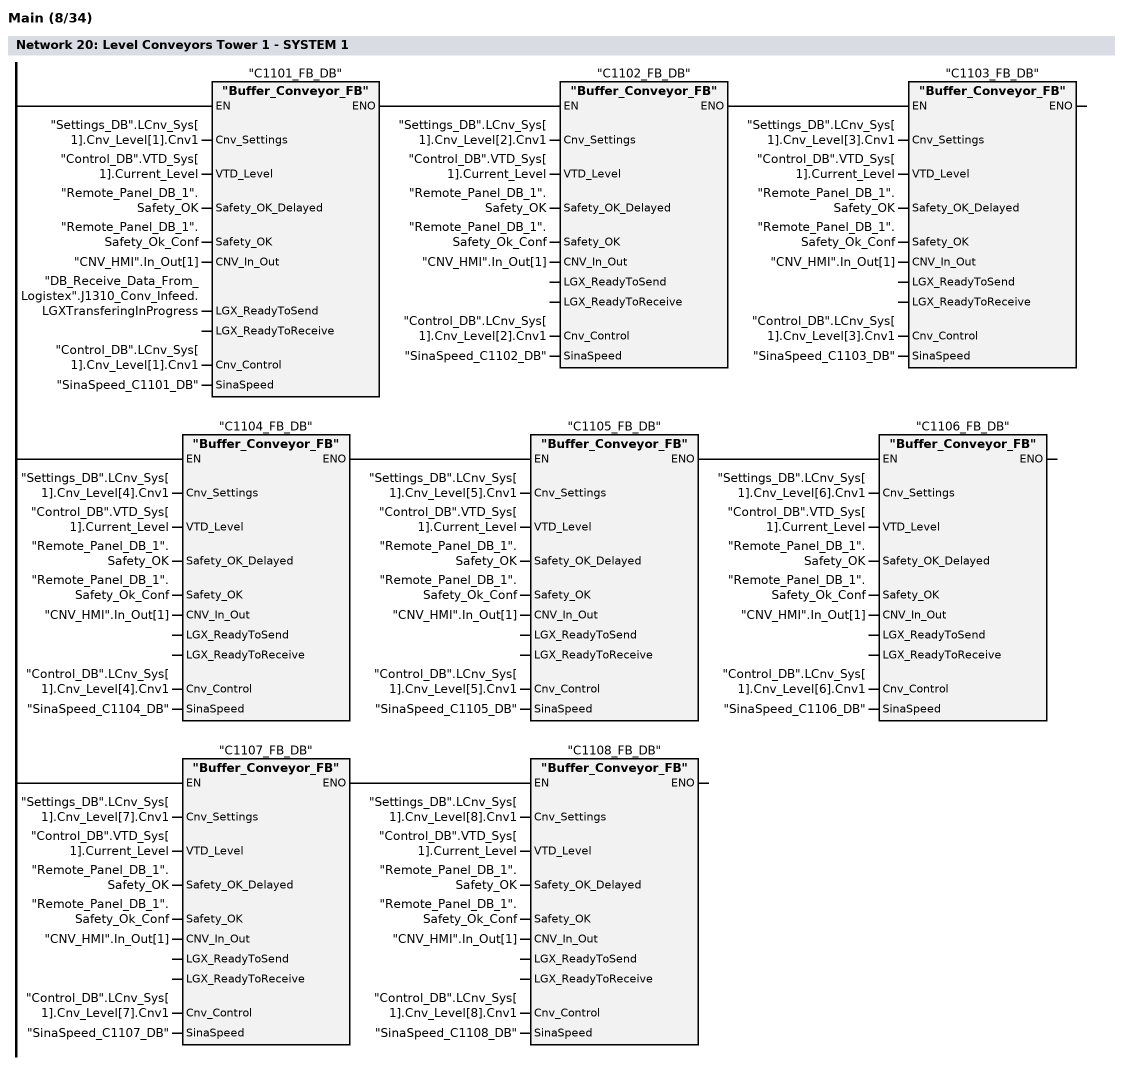
   RUNG wire#powerrail
      "C1101_FB_DB"(Cnv_Settings := "Settings_DB".LCnv_Sys[1].Cnv_Level[1].Cnv1, VTD_Level := "Control_DB".VTD_Sys[1].Current_Level, Safety_OK_Delayed := "Remote_Panel_DB_1".Safety_OK, Safety_OK := "Remote_Panel_DB_1".Safety_Ok_Conf, CNV_In_Out := "CNV_HMI".In_Out[1], LGX_ReadyToSend := "DB_Receive_Data_From_Logistex".J1310_Conv_Infeed.LGXTransferingInProgress, LGX_ReadyToReceive :=, Cnv_Control := "Control_DB".LCnv_Sys[1].Cnv_Level[1].Cnv1, SinaSpeed := "SinaSpeed_C1101_DB")
      "C1102_FB_DB"(Cnv_Settings := "Settings_DB".LCnv_Sys[1].Cnv_Level[2].Cnv1, VTD_Level := "Control_DB".VTD_Sys[1].Current_Level, Safety_OK_Delayed := "Remote_Panel_DB_1".Safety_OK, Safety_OK := "Remote_Panel_DB_1".Safety_Ok_Conf, CNV_In_Out := "CNV_HMI".In_Out[1], LGX_ReadyToSend :=, LGX_ReadyToReceive :=, Cnv_Control := "Control_DB".LCnv_Sys[1].Cnv_Level[2].Cnv1, SinaSpeed := "SinaSpeed_C1102_DB")
      "C1103_FB_DB"(Cnv_Settings := "Settings_DB".LCnv_Sys[1].Cnv_Level[3].Cnv1, VTD_Level := "Control_DB".VTD_Sys[1].Current_Level, Safety_OK_Delayed := "Remote_Panel_DB_1".Safety_OK, Safety_OK := "Remote_Panel_DB_1".Safety_Ok_Conf, CNV_In_Out := "CNV_HMI".In_Out[1], LGX_ReadyToSend :=, LGX_ReadyToReceive :=, Cnv_Control := "Control_DB".LCnv_Sys[1].Cnv_Level[3].Cnv1, SinaSpeed := "SinaSpeed_C1103_DB")
   END_RUNG
   RUNG wire#powerrail
      "C1104_FB_DB"(Cnv_Settings := "Settings_DB".LCnv_Sys[1].Cnv_Level[4].Cnv1, VTD_Level := "Control_DB".VTD_Sys[1].Current_Level, Safety_OK_Delayed := "Remote_Panel_DB_1".Safety_OK, Safety_OK := "Remote_Panel_DB_1".Safety_Ok_Conf, CNV_In_Out := "CNV_HMI".In_Out[1], LGX_ReadyToSend :=, LGX_ReadyToReceive :=, Cnv_Control := "Control_DB".LCnv_Sys[1].Cnv_Level[4].Cnv1, SinaSpeed := "SinaSpeed_C1104_DB")
      "C1105_FB_DB"(Cnv_Settings := "Settings_DB".LCnv_Sys[1].Cnv_Level[5].Cnv1, VTD_Level := "Control_DB".VTD_Sys[1].Current_Level, Safety_OK_Delayed := "Remote_Panel_DB_1".Safety_OK, Safety_OK := "Remote_Panel_DB_1".Safety_Ok_Conf, CNV_In_Out := "CNV_HMI".In_Out[1], LGX_ReadyToSend :=, LGX_ReadyToReceive :=, Cnv_Control := "Control_DB".LCnv_Sys[1].Cnv_Level[5].Cnv1, SinaSpeed := "SinaSpeed_C1105_DB")
      "C1106_FB_DB"(Cnv_Settings := "Settings_DB".LCnv_Sys[1].Cnv_Level[6].Cnv1, VTD_Level := "Control_DB".VTD_Sys[1].Current_Level, Safety_OK_Delayed := "Remote_Panel_DB_1".Safety_OK, Safety_OK := "Remote_Panel_DB_1".Safety_Ok_Conf, CNV_In_Out := "CNV_HMI".In_Out[1], LGX_ReadyToSend :=, LGX_ReadyToReceive :=, Cnv_Control := "Control_DB".LCnv_Sys[1].Cnv_Level[6].Cnv1, SinaSpeed := "SinaSpeed_C1106_DB")
   END_RUNG
   RUNG wire#powerrail
      "C1107_FB_DB"(Cnv_Settings := "Settings_DB".LCnv_Sys[1].Cnv_Level[7].Cnv1, VTD_Level := "Control_DB".VTD_Sys[1].Current_Level, Safety_OK_Delayed := "Remote_Panel_DB_1".Safety_OK, Safety_OK := "Remote_Panel_DB_1".Safety_Ok_Conf, CNV_In_Out := "CNV_HMI".In_Out[1], LGX_ReadyToSend :=, LGX_ReadyToReceive :=, Cnv_Control := "Control_DB".LCnv_Sys[1].Cnv_Level[7].Cnv1, SinaSpeed := "SinaSpeed_C1107_DB")
      "C1108_FB_DB"(Cnv_Settings := "Settings_DB".LCnv_Sys[1].Cnv_Level[8].Cnv1, VTD_Level := "Control_DB".VTD_Sys[1].Current_Level, Safety_OK_Delayed := "Remote_Panel_DB_1".Safety_OK, Safety_OK := "Remote_Panel_DB_1".Safety_Ok_Conf, CNV_In_Out := "CNV_HMI".In_Out[1], LGX_ReadyToSend :=, LGX_ReadyToReceive :=, Cnv_Control := "Control_DB".LCnv_Sys[1].Cnv_Level[8].Cnv1, SinaSpeed := "SinaSpeed_C1108_DB")
   END_RUNG
   // the same network as SCL:
   "C1101_FB_DB"(Cnv_Settings := "Settings_DB".LCnv_Sys[1].Cnv_Level[1].Cnv1,   // "Buffer_Conveyor_FB"
                 VTD_Level := "Control_DB".VTD_Sys[1].Current_Level,
                 Safety_OK_Delayed := "Remote_Panel_DB_1".Safety_OK,
                 Safety_OK := "Remote_Panel_DB_1".Safety_Ok_Conf,
                 CNV_In_Out := "CNV_HMI".In_Out[1],
                 LGX_ReadyToSend := "DB_Receive_Data_From_Logistex".J1310_Conv_Infeed.LGXTransferingInProgress,
                 Cnv_Control := "Control_DB".LCnv_Sys[1].Cnv_Level[1].Cnv1,
                 SinaSpeed := "SinaSpeed_C1101_DB",
                 ENO => #_w1);
   "C1102_FB_DB"(EN := #_w1,   // "Buffer_Conveyor_FB"
                 Cnv_Settings := "Settings_DB".LCnv_Sys[1].Cnv_Level[2].Cnv1,
                 VTD_Level := "Control_DB".VTD_Sys[1].Current_Level,
                 Safety_OK_Delayed := "Remote_Panel_DB_1".Safety_OK,
                 Safety_OK := "Remote_Panel_DB_1".Safety_Ok_Conf,
                 CNV_In_Out := "CNV_HMI".In_Out[1],
                 Cnv_Control := "Control_DB".LCnv_Sys[1].Cnv_Level[2].Cnv1,
                 SinaSpeed := "SinaSpeed_C1102_DB",
                 ENO => #_w2);
   IF #_w2 THEN
       "C1103_FB_DB"(Cnv_Settings := "Settings_DB".LCnv_Sys[1].Cnv_Level[3].Cnv1,   // "Buffer_Conveyor_FB"
                     VTD_Level := "Control_DB".VTD_Sys[1].Current_Level,
                     Safety_OK_Delayed := "Remote_Panel_DB_1".Safety_OK,
                     Safety_OK := "Remote_Panel_DB_1".Safety_Ok_Conf,
                     CNV_In_Out := "CNV_HMI".In_Out[1],
                     Cnv_Control := "Control_DB".LCnv_Sys[1].Cnv_Level[3].Cnv1,
                     SinaSpeed := "SinaSpeed_C1103_DB");
   END_IF;
   "C1104_FB_DB"(Cnv_Settings := "Settings_DB".LCnv_Sys[1].Cnv_Level[4].Cnv1,   // "Buffer_Conveyor_FB"
                 VTD_Level := "Control_DB".VTD_Sys[1].Current_Level,
                 Safety_OK_Delayed := "Remote_Panel_DB_1".Safety_OK,
                 Safety_OK := "Remote_Panel_DB_1".Safety_Ok_Conf,
                 CNV_In_Out := "CNV_HMI".In_Out[1],
                 Cnv_Control := "Control_DB".LCnv_Sys[1].Cnv_Level[4].Cnv1,
                 SinaSpeed := "SinaSpeed_C1104_DB",
                 ENO => #_w3);
   "C1105_FB_DB"(EN := #_w3,   // "Buffer_Conveyor_FB"
                 Cnv_Settings := "Settings_DB".LCnv_Sys[1].Cnv_Level[5].Cnv1,
                 VTD_Level := "Control_DB".VTD_Sys[1].Current_Level,
                 Safety_OK_Delayed := "Remote_Panel_DB_1".Safety_OK,
                 Safety_OK := "Remote_Panel_DB_1".Safety_Ok_Conf,
                 CNV_In_Out := "CNV_HMI".In_Out[1],
                 Cnv_Control := "Control_DB".LCnv_Sys[1].Cnv_Level[5].Cnv1,
                 SinaSpeed := "SinaSpeed_C1105_DB",
                 ENO => #_w4);
   IF #_w4 THEN
       "C1106_FB_DB"(Cnv_Settings := "Settings_DB".LCnv_Sys[1].Cnv_Level[6].Cnv1,   // "Buffer_Conveyor_FB"
                     VTD_Level := "Control_DB".VTD_Sys[1].Current_Level,
                     Safety_OK_Delayed := "Remote_Panel_DB_1".Safety_OK,
                     Safety_OK := "Remote_Panel_DB_1".Safety_Ok_Conf,
                     CNV_In_Out := "CNV_HMI".In_Out[1],
                     Cnv_Control := "Control_DB".LCnv_Sys[1].Cnv_Level[6].Cnv1,
                     SinaSpeed := "SinaSpeed_C1106_DB");
   END_IF;
   "C1107_FB_DB"(Cnv_Settings := "Settings_DB".LCnv_Sys[1].Cnv_Level[7].Cnv1,   // "Buffer_Conveyor_FB"
                 VTD_Level := "Control_DB".VTD_Sys[1].Current_Level,
                 Safety_OK_Delayed := "Remote_Panel_DB_1".Safety_OK,
                 Safety_OK := "Remote_Panel_DB_1".Safety_Ok_Conf,
                 CNV_In_Out := "CNV_HMI".In_Out[1],
                 Cnv_Control := "Control_DB".LCnv_Sys[1].Cnv_Level[7].Cnv1,
                 SinaSpeed := "SinaSpeed_C1107_DB",
                 ENO => #_w5);
   IF #_w5 THEN
       "C1108_FB_DB"(Cnv_Settings := "Settings_DB".LCnv_Sys[1].Cnv_Level[8].Cnv1,   // "Buffer_Conveyor_FB"
                     VTD_Level := "Control_DB".VTD_Sys[1].Current_Level,
                     Safety_OK_Delayed := "Remote_Panel_DB_1".Safety_OK,
                     Safety_OK := "Remote_Panel_DB_1".Safety_Ok_Conf,
                     CNV_In_Out := "CNV_HMI".In_Out[1],
                     Cnv_Control := "Control_DB".LCnv_Sys[1].Cnv_Level[8].Cnv1,
                     SinaSpeed := "SinaSpeed_C1108_DB");
   END_IF;
END_REGION

REGION Network 21: Level Conveyors Tower 2 - SYSTEM 1
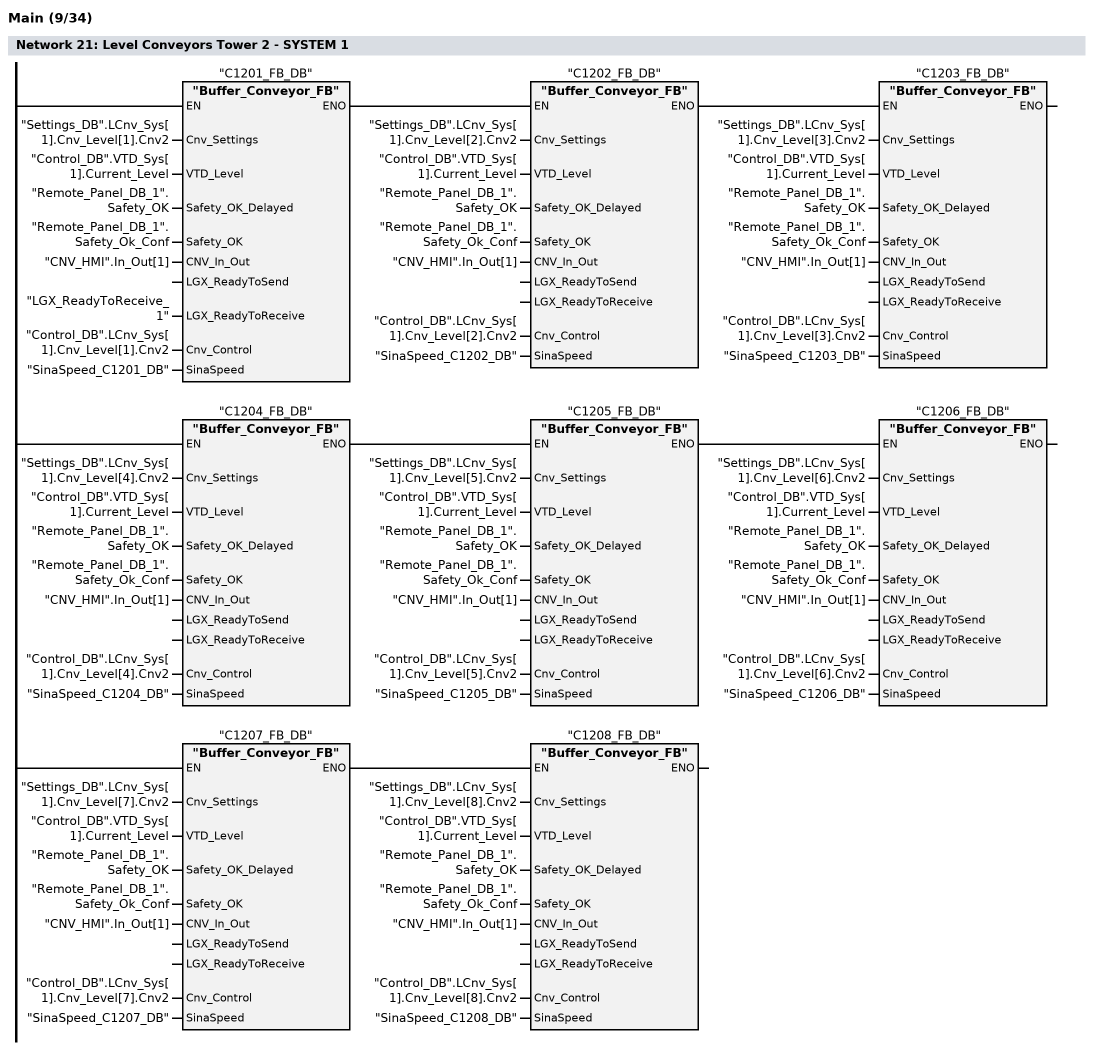
   RUNG wire#powerrail
      "C1201_FB_DB"(Cnv_Settings := "Settings_DB".LCnv_Sys[1].Cnv_Level[1].Cnv2, VTD_Level := "Control_DB".VTD_Sys[1].Current_Level, Safety_OK_Delayed := "Remote_Panel_DB_1".Safety_OK, Safety_OK := "Remote_Panel_DB_1".Safety_Ok_Conf, CNV_In_Out := "CNV_HMI".In_Out[1], LGX_ReadyToSend :=, LGX_ReadyToReceive := "LGX_ReadyToReceive_1", Cnv_Control := "Control_DB".LCnv_Sys[1].Cnv_Level[1].Cnv2, SinaSpeed := "SinaSpeed_C1201_DB")
      "C1202_FB_DB"(Cnv_Settings := "Settings_DB".LCnv_Sys[1].Cnv_Level[2].Cnv2, VTD_Level := "Control_DB".VTD_Sys[1].Current_Level, Safety_OK_Delayed := "Remote_Panel_DB_1".Safety_OK, Safety_OK := "Remote_Panel_DB_1".Safety_Ok_Conf, CNV_In_Out := "CNV_HMI".In_Out[1], LGX_ReadyToSend :=, LGX_ReadyToReceive :=, Cnv_Control := "Control_DB".LCnv_Sys[1].Cnv_Level[2].Cnv2, SinaSpeed := "SinaSpeed_C1202_DB")
      "C1203_FB_DB"(Cnv_Settings := "Settings_DB".LCnv_Sys[1].Cnv_Level[3].Cnv2, VTD_Level := "Control_DB".VTD_Sys[1].Current_Level, Safety_OK_Delayed := "Remote_Panel_DB_1".Safety_OK, Safety_OK := "Remote_Panel_DB_1".Safety_Ok_Conf, CNV_In_Out := "CNV_HMI".In_Out[1], LGX_ReadyToSend :=, LGX_ReadyToReceive :=, Cnv_Control := "Control_DB".LCnv_Sys[1].Cnv_Level[3].Cnv2, SinaSpeed := "SinaSpeed_C1203_DB")
   END_RUNG
   RUNG wire#powerrail
      "C1204_FB_DB"(Cnv_Settings := "Settings_DB".LCnv_Sys[1].Cnv_Level[4].Cnv2, VTD_Level := "Control_DB".VTD_Sys[1].Current_Level, Safety_OK_Delayed := "Remote_Panel_DB_1".Safety_OK, Safety_OK := "Remote_Panel_DB_1".Safety_Ok_Conf, CNV_In_Out := "CNV_HMI".In_Out[1], LGX_ReadyToSend :=, LGX_ReadyToReceive :=, Cnv_Control := "Control_DB".LCnv_Sys[1].Cnv_Level[4].Cnv2, SinaSpeed := "SinaSpeed_C1204_DB")
      "C1205_FB_DB"(Cnv_Settings := "Settings_DB".LCnv_Sys[1].Cnv_Level[5].Cnv2, VTD_Level := "Control_DB".VTD_Sys[1].Current_Level, Safety_OK_Delayed := "Remote_Panel_DB_1".Safety_OK, Safety_OK := "Remote_Panel_DB_1".Safety_Ok_Conf, CNV_In_Out := "CNV_HMI".In_Out[1], LGX_ReadyToSend :=, LGX_ReadyToReceive :=, Cnv_Control := "Control_DB".LCnv_Sys[1].Cnv_Level[5].Cnv2, SinaSpeed := "SinaSpeed_C1205_DB")
      "C1206_FB_DB"(Cnv_Settings := "Settings_DB".LCnv_Sys[1].Cnv_Level[6].Cnv2, VTD_Level := "Control_DB".VTD_Sys[1].Current_Level, Safety_OK_Delayed := "Remote_Panel_DB_1".Safety_OK, Safety_OK := "Remote_Panel_DB_1".Safety_Ok_Conf, CNV_In_Out := "CNV_HMI".In_Out[1], LGX_ReadyToSend :=, LGX_ReadyToReceive :=, Cnv_Control := "Control_DB".LCnv_Sys[1].Cnv_Level[6].Cnv2, SinaSpeed := "SinaSpeed_C1206_DB")
   END_RUNG
   RUNG wire#powerrail
      "C1207_FB_DB"(Cnv_Settings := "Settings_DB".LCnv_Sys[1].Cnv_Level[7].Cnv2, VTD_Level := "Control_DB".VTD_Sys[1].Current_Level, Safety_OK_Delayed := "Remote_Panel_DB_1".Safety_OK, Safety_OK := "Remote_Panel_DB_1".Safety_Ok_Conf, CNV_In_Out := "CNV_HMI".In_Out[1], LGX_ReadyToSend :=, LGX_ReadyToReceive :=, Cnv_Control := "Control_DB".LCnv_Sys[1].Cnv_Level[7].Cnv2, SinaSpeed := "SinaSpeed_C1207_DB")
      "C1208_FB_DB"(Cnv_Settings := "Settings_DB".LCnv_Sys[1].Cnv_Level[8].Cnv2, VTD_Level := "Control_DB".VTD_Sys[1].Current_Level, Safety_OK_Delayed := "Remote_Panel_DB_1".Safety_OK, Safety_OK := "Remote_Panel_DB_1".Safety_Ok_Conf, CNV_In_Out := "CNV_HMI".In_Out[1], LGX_ReadyToSend :=, LGX_ReadyToReceive :=, Cnv_Control := "Control_DB".LCnv_Sys[1].Cnv_Level[8].Cnv2, SinaSpeed := "SinaSpeed_C1208_DB")
   END_RUNG
   // the same network as SCL:
   "C1201_FB_DB"(Cnv_Settings := "Settings_DB".LCnv_Sys[1].Cnv_Level[1].Cnv2,   // "Buffer_Conveyor_FB"
                 VTD_Level := "Control_DB".VTD_Sys[1].Current_Level,
                 Safety_OK_Delayed := "Remote_Panel_DB_1".Safety_OK,
                 Safety_OK := "Remote_Panel_DB_1".Safety_Ok_Conf,
                 CNV_In_Out := "CNV_HMI".In_Out[1],
                 LGX_ReadyToReceive := "LGX_ReadyToReceive_1",
                 Cnv_Control := "Control_DB".LCnv_Sys[1].Cnv_Level[1].Cnv2,
                 SinaSpeed := "SinaSpeed_C1201_DB",
                 ENO => #_w1);
   "C1202_FB_DB"(EN := #_w1,   // "Buffer_Conveyor_FB"
                 Cnv_Settings := "Settings_DB".LCnv_Sys[1].Cnv_Level[2].Cnv2,
                 VTD_Level := "Control_DB".VTD_Sys[1].Current_Level,
                 Safety_OK_Delayed := "Remote_Panel_DB_1".Safety_OK,
                 Safety_OK := "Remote_Panel_DB_1".Safety_Ok_Conf,
                 CNV_In_Out := "CNV_HMI".In_Out[1],
                 Cnv_Control := "Control_DB".LCnv_Sys[1].Cnv_Level[2].Cnv2,
                 SinaSpeed := "SinaSpeed_C1202_DB",
                 ENO => #_w2);
   IF #_w2 THEN
       "C1203_FB_DB"(Cnv_Settings := "Settings_DB".LCnv_Sys[1].Cnv_Level[3].Cnv2,   // "Buffer_Conveyor_FB"
                     VTD_Level := "Control_DB".VTD_Sys[1].Current_Level,
                     Safety_OK_Delayed := "Remote_Panel_DB_1".Safety_OK,
                     Safety_OK := "Remote_Panel_DB_1".Safety_Ok_Conf,
                     CNV_In_Out := "CNV_HMI".In_Out[1],
                     Cnv_Control := "Control_DB".LCnv_Sys[1].Cnv_Level[3].Cnv2,
                     SinaSpeed := "SinaSpeed_C1203_DB");
   END_IF;
   "C1204_FB_DB"(Cnv_Settings := "Settings_DB".LCnv_Sys[1].Cnv_Level[4].Cnv2,   // "Buffer_Conveyor_FB"
                 VTD_Level := "Control_DB".VTD_Sys[1].Current_Level,
                 Safety_OK_Delayed := "Remote_Panel_DB_1".Safety_OK,
                 Safety_OK := "Remote_Panel_DB_1".Safety_Ok_Conf,
                 CNV_In_Out := "CNV_HMI".In_Out[1],
                 Cnv_Control := "Control_DB".LCnv_Sys[1].Cnv_Level[4].Cnv2,
                 SinaSpeed := "SinaSpeed_C1204_DB",
                 ENO => #_w3);
   "C1205_FB_DB"(EN := #_w3,   // "Buffer_Conveyor_FB"
                 Cnv_Settings := "Settings_DB".LCnv_Sys[1].Cnv_Level[5].Cnv2,
                 VTD_Level := "Control_DB".VTD_Sys[1].Current_Level,
                 Safety_OK_Delayed := "Remote_Panel_DB_1".Safety_OK,
                 Safety_OK := "Remote_Panel_DB_1".Safety_Ok_Conf,
                 CNV_In_Out := "CNV_HMI".In_Out[1],
                 Cnv_Control := "Control_DB".LCnv_Sys[1].Cnv_Level[5].Cnv2,
                 SinaSpeed := "SinaSpeed_C1205_DB",
                 ENO => #_w4);
   IF #_w4 THEN
       "C1206_FB_DB"(Cnv_Settings := "Settings_DB".LCnv_Sys[1].Cnv_Level[6].Cnv2,   // "Buffer_Conveyor_FB"
                     VTD_Level := "Control_DB".VTD_Sys[1].Current_Level,
                     Safety_OK_Delayed := "Remote_Panel_DB_1".Safety_OK,
                     Safety_OK := "Remote_Panel_DB_1".Safety_Ok_Conf,
                     CNV_In_Out := "CNV_HMI".In_Out[1],
                     Cnv_Control := "Control_DB".LCnv_Sys[1].Cnv_Level[6].Cnv2,
                     SinaSpeed := "SinaSpeed_C1206_DB");
   END_IF;
   "C1207_FB_DB"(Cnv_Settings := "Settings_DB".LCnv_Sys[1].Cnv_Level[7].Cnv2,   // "Buffer_Conveyor_FB"
                 VTD_Level := "Control_DB".VTD_Sys[1].Current_Level,
                 Safety_OK_Delayed := "Remote_Panel_DB_1".Safety_OK,
                 Safety_OK := "Remote_Panel_DB_1".Safety_Ok_Conf,
                 CNV_In_Out := "CNV_HMI".In_Out[1],
                 Cnv_Control := "Control_DB".LCnv_Sys[1].Cnv_Level[7].Cnv2,
                 SinaSpeed := "SinaSpeed_C1207_DB",
                 ENO => #_w5);
   IF #_w5 THEN
       "C1208_FB_DB"(Cnv_Settings := "Settings_DB".LCnv_Sys[1].Cnv_Level[8].Cnv2,   // "Buffer_Conveyor_FB"
                     VTD_Level := "Control_DB".VTD_Sys[1].Current_Level,
                     Safety_OK_Delayed := "Remote_Panel_DB_1".Safety_OK,
                     Safety_OK := "Remote_Panel_DB_1".Safety_Ok_Conf,
                     CNV_In_Out := "CNV_HMI".In_Out[1],
                     Cnv_Control := "Control_DB".LCnv_Sys[1].Cnv_Level[8].Cnv2,
                     SinaSpeed := "SinaSpeed_C1208_DB");
   END_IF;
END_REGION

REGION Network 22: SAFETY STOPPERS Tower 1 - SYSTEM 1
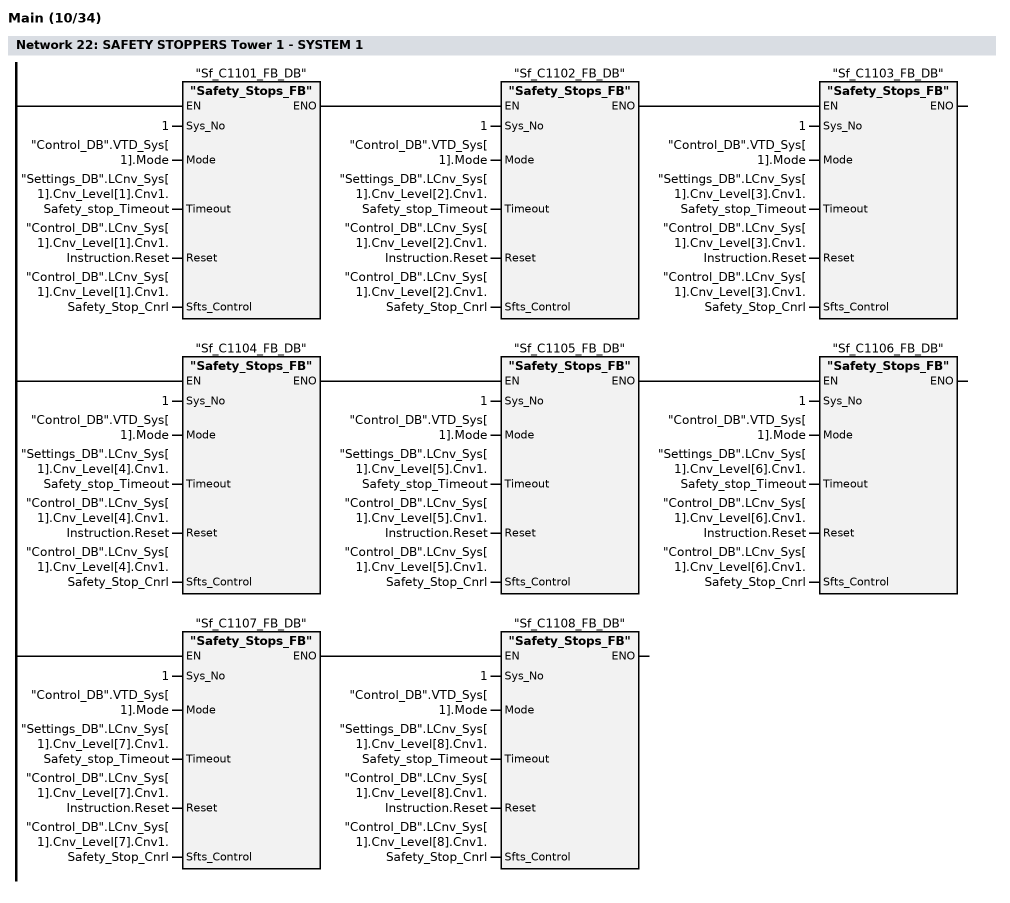
   RUNG wire#powerrail
      "Sf_C1101_FB_DB"(Sys_No := 1, Mode := "Control_DB".VTD_Sys[1].Mode, Timeout := "Settings_DB".LCnv_Sys[1].Cnv_Level[1].Cnv1.Safety_stop_Timeout, Reset := "Control_DB".LCnv_Sys[1].Cnv_Level[1].Cnv1.Instruction.Reset, Sfts_Control := "Control_DB".LCnv_Sys[1].Cnv_Level[1].Cnv1.Safety_Stop_Cnrl)
      "Sf_C1102_FB_DB"(Sys_No := 1, Mode := "Control_DB".VTD_Sys[1].Mode, Timeout := "Settings_DB".LCnv_Sys[1].Cnv_Level[2].Cnv1.Safety_stop_Timeout, Reset := "Control_DB".LCnv_Sys[1].Cnv_Level[2].Cnv1.Instruction.Reset, Sfts_Control := "Control_DB".LCnv_Sys[1].Cnv_Level[2].Cnv1.Safety_Stop_Cnrl)
      "Sf_C1103_FB_DB"(Sys_No := 1, Mode := "Control_DB".VTD_Sys[1].Mode, Timeout := "Settings_DB".LCnv_Sys[1].Cnv_Level[3].Cnv1.Safety_stop_Timeout, Reset := "Control_DB".LCnv_Sys[1].Cnv_Level[3].Cnv1.Instruction.Reset, Sfts_Control := "Control_DB".LCnv_Sys[1].Cnv_Level[3].Cnv1.Safety_Stop_Cnrl)
   END_RUNG
   RUNG wire#powerrail
      "Sf_C1104_FB_DB"(Sys_No := 1, Mode := "Control_DB".VTD_Sys[1].Mode, Timeout := "Settings_DB".LCnv_Sys[1].Cnv_Level[4].Cnv1.Safety_stop_Timeout, Reset := "Control_DB".LCnv_Sys[1].Cnv_Level[4].Cnv1.Instruction.Reset, Sfts_Control := "Control_DB".LCnv_Sys[1].Cnv_Level[4].Cnv1.Safety_Stop_Cnrl)
      "Sf_C1105_FB_DB"(Sys_No := 1, Mode := "Control_DB".VTD_Sys[1].Mode, Timeout := "Settings_DB".LCnv_Sys[1].Cnv_Level[5].Cnv1.Safety_stop_Timeout, Reset := "Control_DB".LCnv_Sys[1].Cnv_Level[5].Cnv1.Instruction.Reset, Sfts_Control := "Control_DB".LCnv_Sys[1].Cnv_Level[5].Cnv1.Safety_Stop_Cnrl)
      "Sf_C1106_FB_DB"(Sys_No := 1, Mode := "Control_DB".VTD_Sys[1].Mode, Timeout := "Settings_DB".LCnv_Sys[1].Cnv_Level[6].Cnv1.Safety_stop_Timeout, Reset := "Control_DB".LCnv_Sys[1].Cnv_Level[6].Cnv1.Instruction.Reset, Sfts_Control := "Control_DB".LCnv_Sys[1].Cnv_Level[6].Cnv1.Safety_Stop_Cnrl)
   END_RUNG
   RUNG wire#powerrail
      "Sf_C1107_FB_DB"(Sys_No := 1, Mode := "Control_DB".VTD_Sys[1].Mode, Timeout := "Settings_DB".LCnv_Sys[1].Cnv_Level[7].Cnv1.Safety_stop_Timeout, Reset := "Control_DB".LCnv_Sys[1].Cnv_Level[7].Cnv1.Instruction.Reset, Sfts_Control := "Control_DB".LCnv_Sys[1].Cnv_Level[7].Cnv1.Safety_Stop_Cnrl)
      "Sf_C1108_FB_DB"(Sys_No := 1, Mode := "Control_DB".VTD_Sys[1].Mode, Timeout := "Settings_DB".LCnv_Sys[1].Cnv_Level[8].Cnv1.Safety_stop_Timeout, Reset := "Control_DB".LCnv_Sys[1].Cnv_Level[8].Cnv1.Instruction.Reset, Sfts_Control := "Control_DB".LCnv_Sys[1].Cnv_Level[8].Cnv1.Safety_Stop_Cnrl)
   END_RUNG
   // the same network as SCL:
   "Sf_C1101_FB_DB"(Sys_No := 1,   // "Safety_Stops_FB"
                    Mode := "Control_DB".VTD_Sys[1].Mode,
                    Timeout := "Settings_DB".LCnv_Sys[1].Cnv_Level[1].Cnv1.Safety_stop_Timeout,
                    Reset := "Control_DB".LCnv_Sys[1].Cnv_Level[1].Cnv1.Instruction.Reset,
                    Sfts_Control := "Control_DB".LCnv_Sys[1].Cnv_Level[1].Cnv1.Safety_Stop_Cnrl,
                    ENO => #_w1);
   "Sf_C1102_FB_DB"(EN := #_w1,   // "Safety_Stops_FB"
                    Sys_No := 1,
                    Mode := "Control_DB".VTD_Sys[1].Mode,
                    Timeout := "Settings_DB".LCnv_Sys[1].Cnv_Level[2].Cnv1.Safety_stop_Timeout,
                    Reset := "Control_DB".LCnv_Sys[1].Cnv_Level[2].Cnv1.Instruction.Reset,
                    Sfts_Control := "Control_DB".LCnv_Sys[1].Cnv_Level[2].Cnv1.Safety_Stop_Cnrl,
                    ENO => #_w2);
   IF #_w2 THEN
       "Sf_C1103_FB_DB"(Sys_No := 1,   // "Safety_Stops_FB"
                        Mode := "Control_DB".VTD_Sys[1].Mode,
                        Timeout := "Settings_DB".LCnv_Sys[1].Cnv_Level[3].Cnv1.Safety_stop_Timeout,
                        Reset := "Control_DB".LCnv_Sys[1].Cnv_Level[3].Cnv1.Instruction.Reset,
                        Sfts_Control := "Control_DB".LCnv_Sys[1].Cnv_Level[3].Cnv1.Safety_Stop_Cnrl);
   END_IF;
   "Sf_C1104_FB_DB"(Sys_No := 1,   // "Safety_Stops_FB"
                    Mode := "Control_DB".VTD_Sys[1].Mode,
                    Timeout := "Settings_DB".LCnv_Sys[1].Cnv_Level[4].Cnv1.Safety_stop_Timeout,
                    Reset := "Control_DB".LCnv_Sys[1].Cnv_Level[4].Cnv1.Instruction.Reset,
                    Sfts_Control := "Control_DB".LCnv_Sys[1].Cnv_Level[4].Cnv1.Safety_Stop_Cnrl,
                    ENO => #_w3);
   "Sf_C1105_FB_DB"(EN := #_w3,   // "Safety_Stops_FB"
                    Sys_No := 1,
                    Mode := "Control_DB".VTD_Sys[1].Mode,
                    Timeout := "Settings_DB".LCnv_Sys[1].Cnv_Level[5].Cnv1.Safety_stop_Timeout,
                    Reset := "Control_DB".LCnv_Sys[1].Cnv_Level[5].Cnv1.Instruction.Reset,
                    Sfts_Control := "Control_DB".LCnv_Sys[1].Cnv_Level[5].Cnv1.Safety_Stop_Cnrl,
                    ENO => #_w4);
   IF #_w4 THEN
       "Sf_C1106_FB_DB"(Sys_No := 1,   // "Safety_Stops_FB"
                        Mode := "Control_DB".VTD_Sys[1].Mode,
                        Timeout := "Settings_DB".LCnv_Sys[1].Cnv_Level[6].Cnv1.Safety_stop_Timeout,
                        Reset := "Control_DB".LCnv_Sys[1].Cnv_Level[6].Cnv1.Instruction.Reset,
                        Sfts_Control := "Control_DB".LCnv_Sys[1].Cnv_Level[6].Cnv1.Safety_Stop_Cnrl);
   END_IF;
   "Sf_C1107_FB_DB"(Sys_No := 1,   // "Safety_Stops_FB"
                    Mode := "Control_DB".VTD_Sys[1].Mode,
                    Timeout := "Settings_DB".LCnv_Sys[1].Cnv_Level[7].Cnv1.Safety_stop_Timeout,
                    Reset := "Control_DB".LCnv_Sys[1].Cnv_Level[7].Cnv1.Instruction.Reset,
                    Sfts_Control := "Control_DB".LCnv_Sys[1].Cnv_Level[7].Cnv1.Safety_Stop_Cnrl,
                    ENO => #_w5);
   IF #_w5 THEN
       "Sf_C1108_FB_DB"(Sys_No := 1,   // "Safety_Stops_FB"
                        Mode := "Control_DB".VTD_Sys[1].Mode,
                        Timeout := "Settings_DB".LCnv_Sys[1].Cnv_Level[8].Cnv1.Safety_stop_Timeout,
                        Reset := "Control_DB".LCnv_Sys[1].Cnv_Level[8].Cnv1.Instruction.Reset,
                        Sfts_Control := "Control_DB".LCnv_Sys[1].Cnv_Level[8].Cnv1.Safety_Stop_Cnrl);
   END_IF;
END_REGION

REGION Network 23: SAFETY STOPPERS Tower 2 - SYSTEM 1
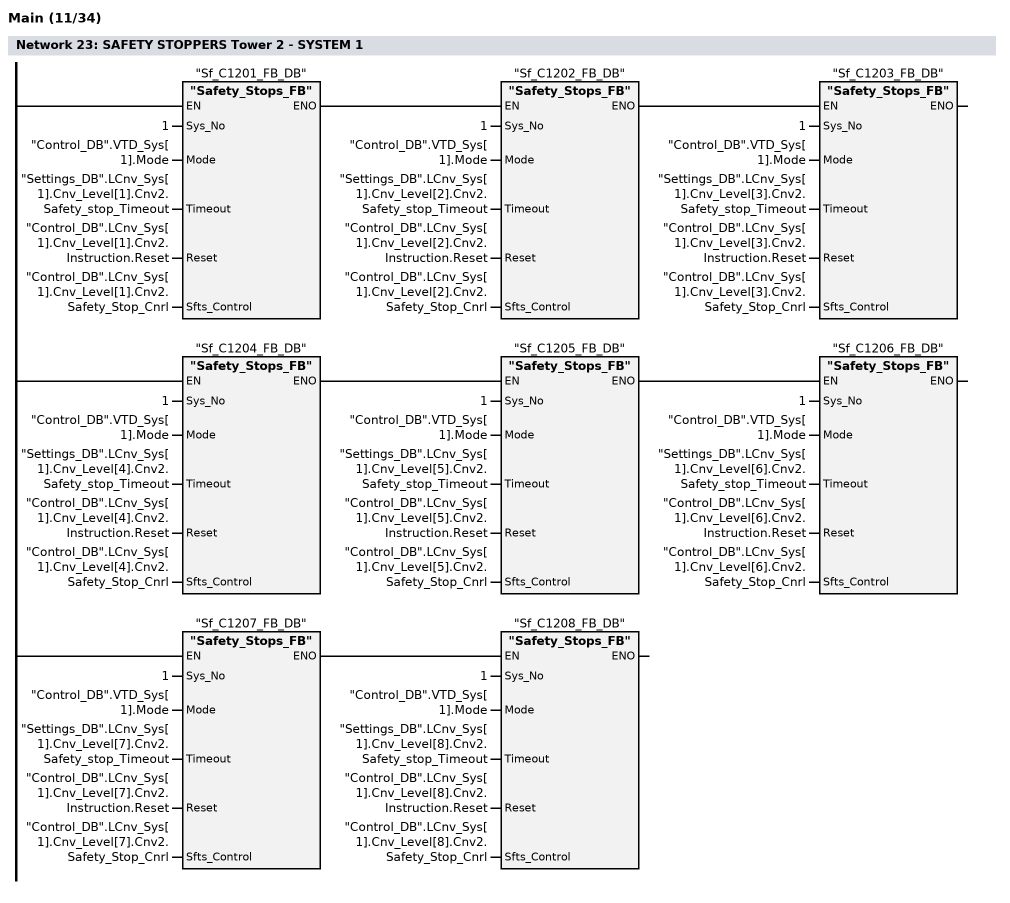
   RUNG wire#powerrail
      "Sf_C1201_FB_DB"(Sys_No := 1, Mode := "Control_DB".VTD_Sys[1].Mode, Timeout := "Settings_DB".LCnv_Sys[1].Cnv_Level[1].Cnv2.Safety_stop_Timeout, Reset := "Control_DB".LCnv_Sys[1].Cnv_Level[1].Cnv2.Instruction.Reset, Sfts_Control := "Control_DB".LCnv_Sys[1].Cnv_Level[1].Cnv2.Safety_Stop_Cnrl)
      "Sf_C1202_FB_DB"(Sys_No := 1, Mode := "Control_DB".VTD_Sys[1].Mode, Timeout := "Settings_DB".LCnv_Sys[1].Cnv_Level[2].Cnv2.Safety_stop_Timeout, Reset := "Control_DB".LCnv_Sys[1].Cnv_Level[2].Cnv2.Instruction.Reset, Sfts_Control := "Control_DB".LCnv_Sys[1].Cnv_Level[2].Cnv2.Safety_Stop_Cnrl)
      "Sf_C1203_FB_DB"(Sys_No := 1, Mode := "Control_DB".VTD_Sys[1].Mode, Timeout := "Settings_DB".LCnv_Sys[1].Cnv_Level[3].Cnv2.Safety_stop_Timeout, Reset := "Control_DB".LCnv_Sys[1].Cnv_Level[3].Cnv2.Instruction.Reset, Sfts_Control := "Control_DB".LCnv_Sys[1].Cnv_Level[3].Cnv2.Safety_Stop_Cnrl)
   END_RUNG
   RUNG wire#powerrail
      "Sf_C1204_FB_DB"(Sys_No := 1, Mode := "Control_DB".VTD_Sys[1].Mode, Timeout := "Settings_DB".LCnv_Sys[1].Cnv_Level[4].Cnv2.Safety_stop_Timeout, Reset := "Control_DB".LCnv_Sys[1].Cnv_Level[4].Cnv2.Instruction.Reset, Sfts_Control := "Control_DB".LCnv_Sys[1].Cnv_Level[4].Cnv2.Safety_Stop_Cnrl)
      "Sf_C1205_FB_DB"(Sys_No := 1, Mode := "Control_DB".VTD_Sys[1].Mode, Timeout := "Settings_DB".LCnv_Sys[1].Cnv_Level[5].Cnv2.Safety_stop_Timeout, Reset := "Control_DB".LCnv_Sys[1].Cnv_Level[5].Cnv2.Instruction.Reset, Sfts_Control := "Control_DB".LCnv_Sys[1].Cnv_Level[5].Cnv2.Safety_Stop_Cnrl)
      "Sf_C1206_FB_DB"(Sys_No := 1, Mode := "Control_DB".VTD_Sys[1].Mode, Timeout := "Settings_DB".LCnv_Sys[1].Cnv_Level[6].Cnv2.Safety_stop_Timeout, Reset := "Control_DB".LCnv_Sys[1].Cnv_Level[6].Cnv2.Instruction.Reset, Sfts_Control := "Control_DB".LCnv_Sys[1].Cnv_Level[6].Cnv2.Safety_Stop_Cnrl)
   END_RUNG
   RUNG wire#powerrail
      "Sf_C1207_FB_DB"(Sys_No := 1, Mode := "Control_DB".VTD_Sys[1].Mode, Timeout := "Settings_DB".LCnv_Sys[1].Cnv_Level[7].Cnv2.Safety_stop_Timeout, Reset := "Control_DB".LCnv_Sys[1].Cnv_Level[7].Cnv2.Instruction.Reset, Sfts_Control := "Control_DB".LCnv_Sys[1].Cnv_Level[7].Cnv2.Safety_Stop_Cnrl)
      "Sf_C1208_FB_DB"(Sys_No := 1, Mode := "Control_DB".VTD_Sys[1].Mode, Timeout := "Settings_DB".LCnv_Sys[1].Cnv_Level[8].Cnv2.Safety_stop_Timeout, Reset := "Control_DB".LCnv_Sys[1].Cnv_Level[8].Cnv2.Instruction.Reset, Sfts_Control := "Control_DB".LCnv_Sys[1].Cnv_Level[8].Cnv2.Safety_Stop_Cnrl)
   END_RUNG
   // the same network as SCL:
   "Sf_C1201_FB_DB"(Sys_No := 1,   // "Safety_Stops_FB"
                    Mode := "Control_DB".VTD_Sys[1].Mode,
                    Timeout := "Settings_DB".LCnv_Sys[1].Cnv_Level[1].Cnv2.Safety_stop_Timeout,
                    Reset := "Control_DB".LCnv_Sys[1].Cnv_Level[1].Cnv2.Instruction.Reset,
                    Sfts_Control := "Control_DB".LCnv_Sys[1].Cnv_Level[1].Cnv2.Safety_Stop_Cnrl,
                    ENO => #_w1);
   "Sf_C1202_FB_DB"(EN := #_w1,   // "Safety_Stops_FB"
                    Sys_No := 1,
                    Mode := "Control_DB".VTD_Sys[1].Mode,
                    Timeout := "Settings_DB".LCnv_Sys[1].Cnv_Level[2].Cnv2.Safety_stop_Timeout,
                    Reset := "Control_DB".LCnv_Sys[1].Cnv_Level[2].Cnv2.Instruction.Reset,
                    Sfts_Control := "Control_DB".LCnv_Sys[1].Cnv_Level[2].Cnv2.Safety_Stop_Cnrl,
                    ENO => #_w2);
   IF #_w2 THEN
       "Sf_C1203_FB_DB"(Sys_No := 1,   // "Safety_Stops_FB"
                        Mode := "Control_DB".VTD_Sys[1].Mode,
                        Timeout := "Settings_DB".LCnv_Sys[1].Cnv_Level[3].Cnv2.Safety_stop_Timeout,
                        Reset := "Control_DB".LCnv_Sys[1].Cnv_Level[3].Cnv2.Instruction.Reset,
                        Sfts_Control := "Control_DB".LCnv_Sys[1].Cnv_Level[3].Cnv2.Safety_Stop_Cnrl);
   END_IF;
   "Sf_C1204_FB_DB"(Sys_No := 1,   // "Safety_Stops_FB"
                    Mode := "Control_DB".VTD_Sys[1].Mode,
                    Timeout := "Settings_DB".LCnv_Sys[1].Cnv_Level[4].Cnv2.Safety_stop_Timeout,
                    Reset := "Control_DB".LCnv_Sys[1].Cnv_Level[4].Cnv2.Instruction.Reset,
                    Sfts_Control := "Control_DB".LCnv_Sys[1].Cnv_Level[4].Cnv2.Safety_Stop_Cnrl,
                    ENO => #_w3);
   "Sf_C1205_FB_DB"(EN := #_w3,   // "Safety_Stops_FB"
                    Sys_No := 1,
                    Mode := "Control_DB".VTD_Sys[1].Mode,
                    Timeout := "Settings_DB".LCnv_Sys[1].Cnv_Level[5].Cnv2.Safety_stop_Timeout,
                    Reset := "Control_DB".LCnv_Sys[1].Cnv_Level[5].Cnv2.Instruction.Reset,
                    Sfts_Control := "Control_DB".LCnv_Sys[1].Cnv_Level[5].Cnv2.Safety_Stop_Cnrl,
                    ENO => #_w4);
   IF #_w4 THEN
       "Sf_C1206_FB_DB"(Sys_No := 1,   // "Safety_Stops_FB"
                        Mode := "Control_DB".VTD_Sys[1].Mode,
                        Timeout := "Settings_DB".LCnv_Sys[1].Cnv_Level[6].Cnv2.Safety_stop_Timeout,
                        Reset := "Control_DB".LCnv_Sys[1].Cnv_Level[6].Cnv2.Instruction.Reset,
                        Sfts_Control := "Control_DB".LCnv_Sys[1].Cnv_Level[6].Cnv2.Safety_Stop_Cnrl);
   END_IF;
   "Sf_C1207_FB_DB"(Sys_No := 1,   // "Safety_Stops_FB"
                    Mode := "Control_DB".VTD_Sys[1].Mode,
                    Timeout := "Settings_DB".LCnv_Sys[1].Cnv_Level[7].Cnv2.Safety_stop_Timeout,
                    Reset := "Control_DB".LCnv_Sys[1].Cnv_Level[7].Cnv2.Instruction.Reset,
                    Sfts_Control := "Control_DB".LCnv_Sys[1].Cnv_Level[7].Cnv2.Safety_Stop_Cnrl,
                    ENO => #_w5);
   IF #_w5 THEN
       "Sf_C1208_FB_DB"(Sys_No := 1,   // "Safety_Stops_FB"
                        Mode := "Control_DB".VTD_Sys[1].Mode,
                        Timeout := "Settings_DB".LCnv_Sys[1].Cnv_Level[8].Cnv2.Safety_stop_Timeout,
                        Reset := "Control_DB".LCnv_Sys[1].Cnv_Level[8].Cnv2.Instruction.Reset,
                        Sfts_Control := "Control_DB".LCnv_Sys[1].Cnv_Level[8].Cnv2.Safety_Stop_Cnrl);
   END_IF;
END_REGION

REGION Network 24: SYSTEM 2
END_REGION

